      (* Pneomatic ->  FB_Piston *)
'2AAx001',   'Error',   'Waiting for Sensor Open at Open command',
'2AAx002',   'Error',   'Waiting for Sensor NotClose at Open command',
'2AAx003',   'Error',   'Waiting for Sensor Close at Close command',
'2AAx004',   'Error',   'Waiting for Sensor NotOpen at Close command',
'2AAx005',   'Error',   'No Status',
'2AAx006',   'Error',   'No Valve Operation',
'2AAx007',   'Error',   'Not synchronized with last auto-cycle command',
'2AAx008',   'Error',   'Sensors Checking',	 
		(*Process elementts*)
'109x000x001',   'Warning',   'Conveyor 5 is full',
'109x000x002',   'Error',     'Conveyor 5 is full and Conveyor 4 is ready to output full stack',

'109x000x003',   'Warning',   'Slices Stack is Too Light',
'109x000x004',   'Error',     'Slices Stack is Too Light',

'109x000x005',   'Warning',   'Slices Stack is Too Heavy',
'109x000x006',   'Error',     'Slices Stack is Too Heavy',
 
'555x000x001',   'Error',     'Hello world from NIV',

'985x000x001',   'Warning',     'X lens Constant velocity did not reach during coating',



(*Niv Section*)
(*Cycle X Curtain*)
(*Cycle X & Y*)
(*Cycle X & Theta)
(*Nozzle Operation*)
(*Cycle X Curtain*)
(*Cycle X Curtain*)*)




''];		
END_VAR

// ---- 01 Instance/06-Visu/g_Common.TcGVL
{attribute 'qualified_only'}
VAR_GLOBAL
	iContent_Main: INT;

END_VAR

// ---- 01 Instance/07-Mode/GVL_OperMode.TcGVL
VAR_GLOBAL

	eLightTowerState: E_LightTowerState;
	eBuzzerMode: E_BuzzerMode;
	bBuzzerMute: BOOL;

	bPauseMachine: BOOL;
	bResumeMachine: BOOL;
	bResetAllCycles: BOOL;
	
	PauseAll: BOOL;
	PauseAllDelayed: BOOL;
	ResumeAll: BOOL;	

	iActErrors							: INT;
	iActMessages						: INT;
	iActWarning							: INT;

	fbMode	: ARRAY[0..E_ModeZone.eLast] OF FB_ModeSelect;
	stMode	: ARRAY[0..E_ModeZone.eLast] OF ST_Mode;
	stOper	: ARRAY[0..E_ModeZone.eLast] OF ST_OperationButtons;
	
	fbLightTower: ARRAY[0..E_SkidZone.eLast] OF FB_LightTower;
	fbLightTower_Control: ARRAY[0..E_SkidZone.eLast] OF FB_LightTower_Control;



	//Operational Modes	
	stModeMain: ST_Mode;
	
	// Operational Buttons
	stOpMain				:ST_OperationButtons;
	stOpNonPause			:ST_OperationButtons;	

END_VAR

// ---- 01 Instance/12 Analog Sensor/g_AnalogSensor.TcGVL
//{attribute 'qualified_only'}
VAR_GLOBAL	
	fbAnalogSensor			: ARRAY[0..E_ASense_Name.last] OF FB_AnalogSensor;
	
	//arAnalogSensorName		: ARRAY[0..E_ASense_Name.last] OF STRING(12);
	
	//arAnalogSensorRawValue	: ARRAY[0..E_ASense_Name.last] OF INT;

	iAnalogSensor_sel		: INT:=1;
	
	arAnalogSensorNameList	: ARRAY[0..E_ASense_Name.last] OF STRING(12);
	eAnalogSensorNameList	: E_ASense_Name;

	
END_VAR
//{attribute 'qualified_only'}
VAR_GLOBAL PERSISTENT
	//stAnalogSensorSetting	: ARRAY[0..E_Pis_Name.last] OF ST_Piston_Setting_Param;
	stAnalogSensor			: ARRAY[0..E_ASense_Name.last] OF ST_AnalogSensor;
END_VAR

VAR_GLOBAL CONSTANT

END_VAR

// ---- 01 Instance/13 Process Control/g_ProcControl.TcGVL
//{attribute 'qualified_only'}
VAR_GLOBAL
	//concentration
	(*stDetergent					:	ST_ProcessControl	;
	pcDetergent					: 	FB_ProcessControl	;	//detergent local
	stDisinfectant				:	ST_ProcessControl	;
	pcDisinfectant				: 	FB_ProcessControl	;	//detergent local
    //temperature
	stTemperature_Deterg			:	ST_ProcessControl	;
	pcTemperature_Deterg			: 	FB_ProcessControl	;	//detergent Client	
	stTemperature_Dis				:	ST_ProcessControl	;
	pcTemperature_Dis				: 	FB_ProcessControl	;//disinfectant local/client
	
	//flow rate
	stFlow_Rate						:	ST_ProcessControl	;//CIP
	pcFlow_Rate						: 	FB_ProcessControl	;//disinfectant local/client
	stFlow_Rate_2					:	ST_ProcessControl	;//CLient CIP //level control 
	pcFlow_Rate_2					: 	FB_ProcessControl	;//disinfectant local/client //level control 
	
	//colar marinade 
	//pressure
	stPressure						:	ST_ProcessControl	;
	pcPressure						: 	FB_ProcessControl	;//CIP //Client	
	*)
	
	///////////////////ARRAYS///////////////////
	arr_fbProcCntrl			:	ARRAY [0..E_ProcessControl_Name.eProcCntrl_Last] OF FB_ProcessControl	;
	arr_ProcCntrl_NameList	:	ARRAY [0..E_ProcessControl_Name.eProcCntrl_Last] OF STRING	;
	eProcCntrl_Name			: E_ProcessControl_Name;
END_VAR
VAR_GLOBAL PERSISTENT
	arr_stProcCntrl			:	ARRAY [0..E_ProcessControl_Name.eProcCntrl_Last] OF ST_ProcessControl	;
END_VAR

// ---- 03 Project/12 TriBlender/g_HMI_Panel.TcGVL
//{attribute 'qualified_only'}
VAR_GLOBAL
	stVisuPLC_To_PLC		AT %MB1000 : ST_VisuPLC_To_PLC;
	stPLC_To_VisuPLC		AT %MB2000 : ST_PLC_To_VisuPLC;
	
	i_stVisuPLC_To_PLC		AT %I* : ST_VisuPLC_To_PLC;
	q_stPLC_To_VisuPLC		AT %Q* : ST_PLC_To_VisuPLC;	
END_VAR

// ---- 03 Project/15 Production Recipes/g_Prod.TcGVL
{attribute 'qualified_only'}
VAR_GLOBAL PERSISTENT
	
	arrRecipeMarinade	: ARRAY[1..cMax_Prod_Recipe] OF ST_Prod_Recipe;
	arrRecipeColor		: ARRAY[1..cMax_Prod_Recipe] OF ST_Prod_Recipe;
	
	iUserSelected_Marinade	: INT;
	iUserSelected_Color		: INT;
	
	fbProdRecipe_Manage	: FB_ProdRecipe_Manage;
	
	listRecipe_Marinade	: ARRAY[1..cMax_Prod_Recipe] OF STRING(30);
	listRecipe_Color	: ARRAY[1..cMax_Prod_Recipe] OF STRING(30);
	
	dtProdTimePicker	: DATE_AND_TIME;
	dtProdTimeMin		: DATE_AND_TIME;
	dtProdTimeMax		: DATE_AND_TIME;



END_VAR
VAR_GLOBAL CONSTANT 
	cMax_Prod_Recipe	: INT:=10;
	cMaxCompInProduct	: USINT:= 10;
END_VAR

// ---- 03 Project/30 IO/gIO.TcGVL
//{attribute 'qualified_only'}
VAR_GLOBAL
	i_EL			AT %I*	: ARRAY[1..27] 		OF ST_EL18x9;
	q_EL			AT %Q*	: ARRAY[1..11] 		OF ST_EL28x9;
	ai_EL			AT %I*	: ARRAY[1..6] 		OF ST_EL3xx8;
	aq_EL			AT %Q*	: ARRAY[1..1] 		OF ST_EL4xx8;

	
	q_Manifold1 	AT %Q*	: ARRAY[1..24] 		OF ST_VTUG;
	q_Manifold2 	AT %Q*	: ARRAY[1..24] 		OF ST_VTUG;
	q_Manifold3 	AT %Q*	: ARRAY[1..24] 		OF ST_VTUG;

	Nidec					: ARRAY[0..E_Pump_List.last] 		OF ST_Nidec;

	
	arSafe			: ARRAY[1..1] OF ST_TwinSAFE;
	bStateSafe		: BOOL;
	bStateSafe_ES1	: BOOL;
	bStateSafe_ES2	: BOOL;
	bStateSafe_ES3	: BOOL;
	bStateSafe_ES4	: BOOL;
	
	fbScaleFactor: ARRAY[0..E_ASense_Name.last] 		OF FB_ScaleFactor;

	
END_VAR

// ---- 03 Project/g_Data.TcGVL
//{attribute 'qualified_only'}
VAR_GLOBAL PERSISTENT
	gCIP_ValvUL			:	ARRAY [1..8,1..6] OF E_Pis_Name	:=[
																E_Pis_Name.V3004,E_Pis_Name.V3017,E_Pis_Name.V3023,E_Pis_Name.e0_not_in_use,E_Pis_Name.e0_not_in_use,E_Pis_Name.e0_not_in_use,
																E_Pis_Name.V3010,E_Pis_Name.V3027,E_Pis_Name.V3028,E_Pis_Name.e0_not_in_use,E_Pis_Name.e0_not_in_use,E_Pis_Name.e0_not_in_use,
																E_Pis_Name.V4034,E_Pis_Name.V4004,E_Pis_Name.V4017,E_Pis_Name.v4023,E_Pis_Name.e0_not_in_use,E_Pis_Name.e0_not_in_use,
																E_Pis_Name.V4033,E_Pis_Name.V4010,E_Pis_Name.V4027,E_Pis_Name.V4028,E_Pis_Name.e0_not_in_use,E_Pis_Name.e0_not_in_use,
																
																E_Pis_Name.V3113,E_Pis_Name.V3004,E_Pis_Name.V3010,E_Pis_Name.V3023,E_Pis_Name.V3028,E_Pis_Name.e0_not_in_use,
																E_Pis_Name.v2114,E_Pis_Name.V4004,E_Pis_Name.V4010,E_Pis_Name.V2116,E_Pis_Name.V4023,E_Pis_Name.V4028,
																E_Pis_Name.V3017,E_Pis_Name.V3027,E_Pis_Name.e0_not_in_use,E_Pis_Name.e0_not_in_use,E_Pis_Name.e0_not_in_use,E_Pis_Name.e0_not_in_use,
																E_Pis_Name.V4017,E_Pis_Name.v4027,E_Pis_Name.V2115,E_Pis_Name.V4034,E_Pis_Name.V4033,E_Pis_Name.e0_not_in_use														
															];	
	gCIP_ValvUL_Seat	:	ARRAY [1..8,1..6] OF BOOL :=[
															0,1,1,0,0,0, // Client 1 eTank_1,
															0,1,1,0,0,0, // Client 2 eTank_2,
															0,0,1,1,0,0, // Client 3 eTank_3,
															0,0,1,1,0,0, // Client 4 eTank_4,
															0,1,1,0,0,0, // Client 5
															0,1,1,0,0,0, // Client 6
															0,0,0,0,0,0, // Client 7
															0,0,0,1,1,0 // Client 8 
														]	;	//0-Low, 1-Up

	fbElement: ARRAY[1..8] OF FB_Element;
	
	fbIntCon_TriB_T1_Marin	: FB_InterConnection;
	fbIntCon_TriB_T2_Marin	: FB_InterConnection;
	fbIntCon_TriB_T3_Color	: FB_InterConnection;
	fbIntCon_TriB_T4_Color	: FB_InterConnection;
	fbIntCon_ProL_T1_Marin	: FB_InterConnection;
	fbIntCon_ProL_T2_Marin	: FB_InterConnection;
	fbIntCon_ProL_T3_Color	: FB_InterConnection;
	fbIntCon_ProL_T4_Color	: FB_InterConnection;
	
	fbTank1					: FB_ProductionTank;
	fbTank2					: FB_ProductionTank;
	fbTank3					: FB_ProductionTank;
	fbTank4					: FB_ProductionTank;

	fbTankTarget_1				: FB_Tank_Target;
	fbTankTarget_2				: FB_Tank_Target;
	fbTankTarget_3				: FB_Tank_Target;
	fbTankTarget_4				: FB_Tank_Target;

	fbLineSource_Marinade		: FB_Line_Source;
	fbTriBlenderSource_Marinade	: FB_Line_Source;
	fbLineSource_Color			: FB_Line_Source;
	fbTriBlenderSource_Color	: FB_Line_Source;
	
	fbLineTarget_Marinade		: FB_Line_Target;
	fbTriBlenderTarget_Marinade	: FB_Line_Target;
	fbLineTarget_Color			: FB_Line_Target;
	fbTriBlenderTarget_Color	: FB_Line_Target;
	
	fbCIP						: FB_CIP;
	
	fbCIP_Source				: FB_CIP_Source;
	fbCIP_Return				: FB_CIP_Return;
	fbCIP_Client				: FB_CIP_Client;
	
	fbCIP_ClientTank_Marinade	: FB_CIP_ClientTank;
	fbCIP_ClientTank_Color		: FB_CIP_ClientTank;

	fbDissolving				: FB_Dissolving;
	fbTriBlender_Select			: FB_TriBlender_Select;
	eTriBlenderUsage	: E_TriBlenderUsage;
	
	eTriBlenderPipe		: E_TriBlenderPipe;
	eTriBlenderPipe_In	: E_TriBlenderPipe;
	eTriBlenderPipe_Out	: E_TriBlenderPipe;

	ePrL_M_Usage		: E_PrLine_M_LineUsage;
	ePrL_C_Usage		: E_PrLine_C_Usage;
	
	//Pumps
	//fbPumpLine_P4001		:	FB_Pump	;
	//fbPumpLine_P3001		:	FB_Pump	;
	//fbPumpTriblender_TB001	:	FB_Pump	;
	
	arCIP_RequestBufer: ARRAY [0..9] OF ST_CIP_Request;

	//stDev			: 	ARRAY[0..E_OwnerDevice.common] OF 	ST_DeviceErrorHandeling;
	//stDev			: 	ARRAY[0..E_OwnerDevice.common] OF 	ST_OperationButtons;
	
	//Valves
	arr_TankValves					:	ARRAY [1..4] OF st_TankValves		;
	arr_LineSourceValves			:	ARRAY [1..4] OF st_LineSourceValves	;
	arr_TriBlenderSourceValves		:	ARRAY [1..4] OF st_LineSourceValves	;
	arr_LineTargetValves			:	ARRAY [1..4] OF st_LineTargetValves	;
	arr_fbTriBlenderTargetValves	:	ARRAY [1..4] OF st_LineTargetValves	;
	
	//Sensors
	(*lvl_Tank_T91	: ST_Tank_Level	;
	lvl_Tank_T92	: ST_Tank_Level	;
	lvl_Tank_T93	: ST_Tank_Level	;
	lvl_Tank_T94	: ST_Tank_Level	;
	
	lvl_Tank_T91_Analog	:	ST_AnalogSignal	;
	lvl_Tank_T92_Analog	:	ST_AnalogSignal	;
	lvl_Tank_T93_Analog	:	ST_AnalogSignal	;
	lvl_Tank_T94_Analog	:	ST_AnalogSignal	;
	
	fbLvl_Tank_T91	:	FB_TankLevel	;
	fbLvl_Tank_T92	:	FB_TankLevel	;
	fbLvl_Tank_T93	:	FB_TankLevel	;
	fbLvl_Tank_T94	:	FB_TankLevel	;
	
	fb_Tank_T91_Sensors	:	FB_TankSensors	;
	fb_Tank_T92_Sensors	:	FB_TankSensors	;
	fb_Tank_T93_Sensors	:	FB_TankSensors	;
	fb_Tank_T94_Sensors	:	FB_TankSensors	;*)
	
	//Heat Exchanger
	fbHeatExchenger	:	FB_HeatExchanger	;
	stHeatExchanger	:	ST_HeatExchanger	;
	
	////////////////////////////////////////////////////////////////
	arrTanksSens	:	ARRAY [0..E_Tank_Name.last] OF FB_TankSensors;
	stTanksSens		:	ARRAY [0..E_Tank_Name.last] OF ST_Tank_Level;
	
	////////////////////////////////////////////////////////////////
	arr_CIP_Param		:	ARRAY [0..E_CIP_Usage.eLocal] OF ST_CIP_Param		;//9-local, 1..8 cleints
	
	//additional variables
	b_CIP_Run	:	BOOL	;
	bDisolvingProcess_Active: BOOL;
	bDisolvingProcess_Done: BOOL;
	
	ExDuration_Default				: TIME:=T#48H;	//Expiration
	ExDuration_Default_Line			: TIME:=T#24H;	//Expiration
	ExDuration_Default_LineStandby	: TIME:=T#2H;	//Expiration

	//arr_ProdTank		:	ARRAY [0..E_Tank_Name.last] OF ST_ProdParams;
	
	//stTriBlender		: ST_TriBlender;		
	//arrProductionComponents	: ARRAY [0..g_Prod.cMaxCompInProduct-1] OF ST_Component;
END_VAR
VAR_GLOBAL CONSTANT
	
END_VAR

// ---- 00 Library/03 SFC/ITF_FB_SFC_Cycle.TcIO
INTERFACE ITF_FB_SFC_Cycle

METHOD m_Set_SFCFlags_Reference : BOOL
VAR_INPUT
END_VAR
END_METHOD

END_INTERFACE

// ---- 01 Instance/04 Recipe/prg_Call_Recipe_Slow.TcPOU
PROGRAM prg_Call_Recipe_Slow
VAR
	i							: INT;
	bFirstScan					: BOOL:= TRUE;
	ton_RecipeReady				: TON;
	
	
	eRecipeName: E_Recipe_Name;

	r_trigAxisPoints_Loaded: R_TRIG;
	ton_WriteLoaded_Points: TON;
	r_trigRecipe3_loaded: R_TRIG;

	bAllRecipesLoaded: BOOL;
	iRecipeSwitchFrameVar: INT;
	bLoadDefForAll: BOOL;
	
	tPath: STRING(80);
END_VAR

act_Set_StoragePath_For_All();
//act_LoadDeafult();

ton_RecipeReady(PT:=T#1S, IN:=GVL_Recipe.stRecipe[1].bInit AND bFirstScan);
IF ton_RecipeReady.Q THEN;
	bFirstScan:=FALSE;
	bLoadDefForAll:=TRUE;
END_IF




(********************  Other Instances Recipes******************************) // 
FOR eRecipeName:=1 TO E_Recipe_Name.R_Piston_Settings DO	
	fbRecipe[eRecipeName](pstRecipe:=ADR(GVL_Recipe.stRecipe[eRecipeName]), 
			bMemoRecipeUpdated:=, 
			sRecipeDef:=TO_STRING(eRecipeName),
			bLoadDefault:=ar_RecipesLoadDefault[eRecipeName],
			bHMI_FrameActive:=iRecipeSwitchFrameVar=eRecipeName-1,//changed
			sRecipesStoragePath:=ar_RecipesStoragePath[eRecipeName]);
END_FOR
(*			
IF (*fbRecipe_1.bMemoRecipeUpdated AND*) 
fbRecipe_2.bMemoRecipeUpdated 
AND fbRecipe_3.bMemoRecipeUpdated 
AND fbRecipe_4.bMemoRecipeUpdated 
AND fbRecipe_5.bMemoRecipeUpdated 
THEN;
	bAllRecipesLoaded:=TRUE;
ELSE;
	bAllRecipesLoaded:=FALSE;
END_IF
*)

ACTION act_LoadDeafult:
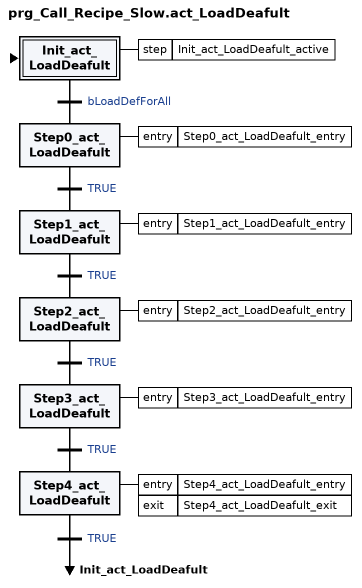
INITIAL_STEP Init_act_LoadDeafult:
    Init_act_LoadDeafult_active(N);  // step action
END_STEP
TRANSITION FROM Init_act_LoadDeafult TO Step0_act_LoadDeafult
    := bLoadDefForAll;
END_TRANSITION
STEP Step0_act_LoadDeafult:  // min time T#2s
    Step0_act_LoadDeafult_entry(P1);  // entry action
END_STEP
TRANSITION FROM Step0_act_LoadDeafult TO Step1_act_LoadDeafult
    := TRUE;
END_TRANSITION
STEP Step1_act_LoadDeafult:  // min time T#2s
    Step1_act_LoadDeafult_entry(P1);  // entry action
END_STEP
TRANSITION FROM Step1_act_LoadDeafult TO Step2_act_LoadDeafult
    := TRUE;
END_TRANSITION
STEP Step2_act_LoadDeafult:  // min time T#2s
    Step2_act_LoadDeafult_entry(P1);  // entry action
END_STEP
TRANSITION FROM Step2_act_LoadDeafult TO Step3_act_LoadDeafult
    := TRUE;
END_TRANSITION
STEP Step3_act_LoadDeafult:  // min time T#2s
    Step3_act_LoadDeafult_entry(P1);  // entry action
END_STEP
TRANSITION FROM Step3_act_LoadDeafult TO Step4_act_LoadDeafult
    := TRUE;
END_TRANSITION
STEP Step4_act_LoadDeafult:  // min time T#2s
    Step4_act_LoadDeafult_entry(P1);  // entry action
    Step4_act_LoadDeafult_exit(P0);  // exit action
END_STEP
TRANSITION FROM Step4_act_LoadDeafult TO Init_act_LoadDeafult
    := TRUE;
END_TRANSITION
END_ACTION

ACTION act_Set_StoragePath_For_All:
FOR eRecipeName:=1 TO E_Recipe_Name.R_Piston_Settings DO;
	GVL_Recipe.ar_RecipesStoragePath_Folder[eRecipeName]:=TO_STRING(eRecipeName);
	tPath:='';
	tPath:=CONCAT(tPath,GVL_Recipe.ar_RecipesStoragePath_Root[GVL_Recipe.eRecipeRootFolder]);
	tPath:=CONCAT(tPath,'\');
	tPath:=CONCAT(tPath,TO_STRING(eRecipeName));
	tPath:=CONCAT(tPath,'\');
	GVL_Recipe.ar_RecipesStoragePath[eRecipeName]:=tPath;
(*
	GVL_Recipe.ar_RecipesStoragePath[eRecipeName]:=
			CONCAT(	GVL_Recipe.ar_RecipesStoragePath_Root[GVL_Recipe.eRecipeRootFolder],'\'); 
	GVL_Recipe.ar_RecipesStoragePath[eRecipeName]:=		
			CONCAT(	GVL_Recipe.ar_RecipesStoragePath[eRecipeName],TO_STRING(eRecipeName));
	GVL_Recipe.ar_RecipesStoragePath[eRecipeName]:=		
			CONCAT(	GVL_Recipe.ar_RecipesStoragePath[eRecipeName],'1');				
	GVL_Recipe.ar_RecipesStoragePath[eRecipeName]:=		
			CONCAT(	GVL_Recipe.ar_RecipesStoragePath[eRecipeName],'\');		
*)	
END_FOR
END_ACTION

ACTION Init_act_LoadDeafult_active:
GVL_Recipe.ar_RecipesLoadDefault[1]:=FALSE;
GVL_Recipe.ar_RecipesLoadDefault[2]:=FALSE;
GVL_Recipe.ar_RecipesLoadDefault[3]:=FALSE;
GVL_Recipe.ar_RecipesLoadDefault[4]:=FALSE;
GVL_Recipe.ar_RecipesLoadDefault[5]:=FALSE;
END_ACTION

ACTION Step0_act_LoadDeafult_entry:
GVL_Recipe.ar_RecipesLoadDefault[1]:=TRUE;
END_ACTION

ACTION Step1_act_LoadDeafult_entry:
GVL_Recipe.ar_RecipesLoadDefault[2]:=TRUE;
END_ACTION

ACTION Step2_act_LoadDeafult_entry:
GVL_Recipe.ar_RecipesLoadDefault[3]:=TRUE;
END_ACTION

ACTION Step3_act_LoadDeafult_entry:
GVL_Recipe.ar_RecipesLoadDefault[4]:=TRUE;
END_ACTION

ACTION Step4_act_LoadDeafult_entry:
GVL_Recipe.ar_RecipesLoadDefault[5]:=TRUE;
END_ACTION

ACTION Step4_act_LoadDeafult_exit:
bLoadDefForAll:=FALSE;
END_ACTION

END_PROGRAM

// ---- POUs/MAIN.TcPOU
PROGRAM MAIN
VAR

	fTotalCIP_Volume: REAL;
	fbWritePersistent: FB_WritePersistentData;
	bTesting		:	BOOL:=FALSE	;
	nI_1			: 	INT		;
	ftg_EStop_Fall	: 	F_TRIG	;
	rs_EStopFall	: 	RS	;
	bTestEstop		:	BOOL:=TRUE	;
	FB_OpenClose_Vlave_4026: FB_OpenClose_Vlave;
	bTemp_Water_Overweight_check: BOOL;
	fbUPS: FB_S_UPS_CX51x0;

	bSetExpeationTime: BOOL;
	i: E_ELEMENT_LIST;
	tExpirationSet_Test: TIME := T#10s;
END_VAR

prg_RealClock();
prg_Piston();
prg_Safety();
prg_MessageManager();
prg_Messages();
prg_Call_OpMode();
prg_IntCheck();
prg_User();
act_ResetPumps();
(*
prg_TriBlender(
		fb_TriBlenderPump:= g_Pump.fbPump[E_Pump_List.TB0001],
		stTriblender:=stTriblender,
		arrComponents:=arrProductionComponents);
*)		
//act_SetAnalogSens_Test();//To be deleted, for testing purposes
act_Call_Sensors_Analog();//To be deleted, for testing purposes
act_Call_Sensors_Analog_1();//To be deleted, for testing purposes
act_Call_ScaleFactor();//To be deleted, for testing purposes
act_Call_ProcessCntrl();

act_SetValves();
act_ClientPump_Select();
act_ClientStirrer_Select();
act_Call_Elements();
act_Call_Elements_Imp();
act_Call_Pumps();
prg_InterCon_Usage();
act_Sensors();
act_HeatExchenger();
act_Call_CIP();
act_Call_Production();

act_Call_For_HMI();

g_SFC.fbSFC_Temp1();

//Temtprary Overweght protection!!!!! DO NOT DELETE
IF fTotalCIP_Volume >=1500 AND FALSE THEN;
	//fbPis[E_Pis_Name.V1022].m_SetByRecipe(stPis:=stPis[E_Pis_Name.V1022], req:=E_Piston_Recipe_State.Release);
	//fbPis[E_Pis_Name.V1019].m_SetByRecipe(stPis:=stPis[E_Pis_Name.V1019], req:=E_Piston_Recipe_State.Release);
	//fbPis[E_Pis_Name.V1016].m_SetByRecipe(stPis:=stPis[E_Pis_Name.V1016], req:=E_Piston_Recipe_State.Release);
	//fbPis[E_Pis_Name.V1011].m_SetByRecipe(stPis:=stPis[E_Pis_Name.V1011], req:=E_Piston_Recipe_State.Release);
	bTemp_Water_Overweight_check:=FALSE;
	fbPrintErrMessageByID(sModuleDescription:='CIP',sActErrorID:='101x000x000');
ELSIF fTotalCIP_Volume < 1480 THEN;
	bTemp_Water_Overweight_check:=TRUE;
END_IF

IF arrTanksSens[E_Tank_Name.T91].get_stTankLevel_OverFlow() THEN;
	fbPis[E_Pis_Name.V1022].m_SetByRecipe(stPis:=stPis[E_Pis_Name.V1022], req:=E_Piston_Recipe_State.Release);
	//print error
	fbPrintErrMessageByID(sModuleDescription:='CIP',sActErrorID:='101x000x001');		
END_IF
IF arrTanksSens[E_Tank_Name.T92].get_stTankLevel_OverFlow() THEN;
	fbPis[E_Pis_Name.V1019].m_SetByRecipe(stPis:=stPis[E_Pis_Name.V1019], req:=E_Piston_Recipe_State.Release);
	//print error
	fbPrintErrMessageByID(sModuleDescription:='CIP',sActErrorID:='101x000x002');		
END_IF
IF arrTanksSens[E_Tank_Name.T93].get_stTankLevel_OverFlow() THEN;
	fbPis[E_Pis_Name.V1016].m_SetByRecipe(stPis:=stPis[E_Pis_Name.V1016], req:=E_Piston_Recipe_State.Release);
	//print error	
	fbPrintErrMessageByID(sModuleDescription:='CIP',sActErrorID:='101x000x003');	
END_IF
IF arrTanksSens[E_Tank_Name.T94].get_stTankLevel_OverFlow() THEN;
	fbPis[E_Pis_Name.V1011].m_SetByRecipe(stPis:=stPis[E_Pis_Name.V1011], req:=E_Piston_Recipe_State.Release);
	//print error
	fbPrintErrMessageByID(sModuleDescription:='CIP',sActErrorID:='101x000x004');		
END_IF
	
IF bSetExpeationTime THEN;
	bSetExpeationTime:=FALSE;
	FOR i:=E_Element_List.eTank_1 TO E_Element_List.eLine_Color DO
		fbElement[i].ExpirationTime:=tExpirationSet_Test;
		
	END_FOR
END_IF
	

mElementList_SetName();

fbWritePersistent(
	NETID:= , 
	PORT:= 851, 
	START:= , 
	TMOUT:= T#3S, 
	MODE:= , 
	BUSY=> , 
	ERR=> , 
	ERRID=> );

fbUPS();

ACTION act_Call_CIP:
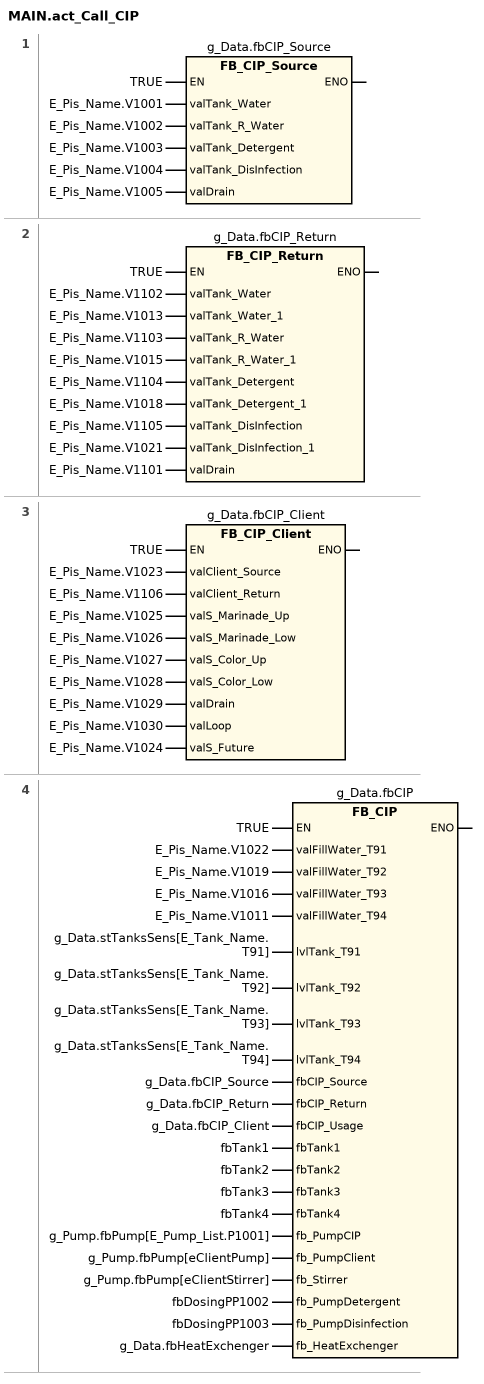
// NETWORK 1
g_Data.fbCIP_Source(
    valTank_Water := E_Pis_Name.V1001,
    valTank_R_Water := E_Pis_Name.V1002,
    valTank_Detergent := E_Pis_Name.V1003,
    valTank_DisInfection := E_Pis_Name.V1004,
    valDrain := E_Pis_Name.V1005); // FB_CIP_Source

// NETWORK 2
g_Data.fbCIP_Return(
    valTank_Water := E_Pis_Name.V1102,
    valTank_Water_1 := E_Pis_Name.V1013,
    valTank_R_Water := E_Pis_Name.V1103,
    valTank_R_Water_1 := E_Pis_Name.V1015,
    valTank_Detergent := E_Pis_Name.V1104,
    valTank_Detergent_1 := E_Pis_Name.V1018,
    valTank_DisInfection := E_Pis_Name.V1105,
    valTank_DisInfection_1 := E_Pis_Name.V1021,
    valDrain := E_Pis_Name.V1101); // FB_CIP_Return

// NETWORK 3
g_Data.fbCIP_Client(
    valClient_Source := E_Pis_Name.V1023,
    valClient_Return := E_Pis_Name.V1106,
    valS_Marinade_Up := E_Pis_Name.V1025,
    valS_Marinade_Low := E_Pis_Name.V1026,
    valS_Color_Up := E_Pis_Name.V1027,
    valS_Color_Low := E_Pis_Name.V1028,
    valDrain := E_Pis_Name.V1029,
    valLoop := E_Pis_Name.V1030,
    valS_Future := E_Pis_Name.V1024); // FB_CIP_Client

// NETWORK 4
g_Data.fbCIP(
    valFillWater_T91 := E_Pis_Name.V1022,
    valFillWater_T92 := E_Pis_Name.V1019,
    valFillWater_T93 := E_Pis_Name.V1016,
    valFillWater_T94 := E_Pis_Name.V1011,
    lvlTank_T91 := g_Data.stTanksSens[E_Tank_Name.T91],
    lvlTank_T92 := g_Data.stTanksSens[E_Tank_Name.T92],
    lvlTank_T93 := g_Data.stTanksSens[E_Tank_Name.T93],
    lvlTank_T94 := g_Data.stTanksSens[E_Tank_Name.T94],
    fbCIP_Source := g_Data.fbCIP_Source,
    fbCIP_Return := g_Data.fbCIP_Return,
    fbCIP_Usage := g_Data.fbCIP_Client,
    fbTank1 := fbTank1,
    fbTank2 := fbTank2,
    fbTank3 := fbTank3,
    fbTank4 := fbTank4,
    fb_PumpCIP := g_Pump.fbPump[E_Pump_List.P1001],
    fb_PumpClient := g_Pump.fbPump[eClientPump],
    fb_Stirrer := g_Pump.fbPump[eClientStirrer],
    fb_PumpDetergent := fbDosingPP1002,
    fb_PumpDisinfection := fbDosingPP1003,
    fb_HeatExchenger := g_Data.fbHeatExchenger); // FB_CIP

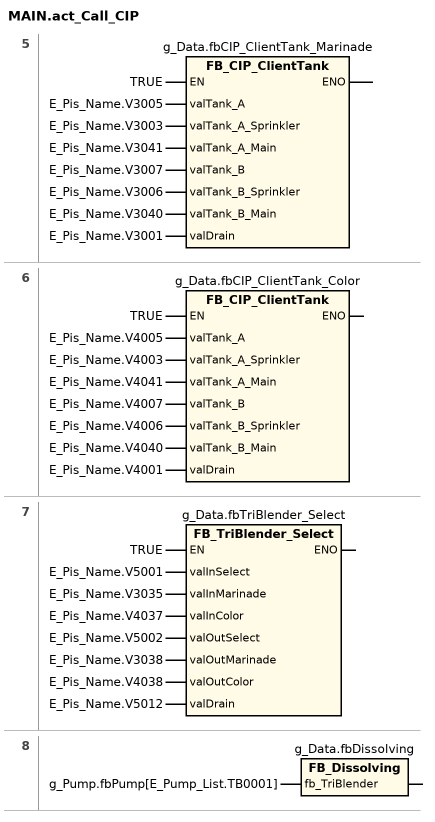
// NETWORK 5
g_Data.fbCIP_ClientTank_Marinade(
    valTank_A := E_Pis_Name.V3005,
    valTank_A_Sprinkler := E_Pis_Name.V3003,
    valTank_A_Main := E_Pis_Name.V3041,
    valTank_B := E_Pis_Name.V3007,
    valTank_B_Sprinkler := E_Pis_Name.V3006,
    valTank_B_Main := E_Pis_Name.V3040,
    valDrain := E_Pis_Name.V3001); // FB_CIP_ClientTank

// NETWORK 6
g_Data.fbCIP_ClientTank_Color(
    valTank_A := E_Pis_Name.V4005,
    valTank_A_Sprinkler := E_Pis_Name.V4003,
    valTank_A_Main := E_Pis_Name.V4041,
    valTank_B := E_Pis_Name.V4007,
    valTank_B_Sprinkler := E_Pis_Name.V4006,
    valTank_B_Main := E_Pis_Name.V4040,
    valDrain := E_Pis_Name.V4001); // FB_CIP_ClientTank

// NETWORK 7
g_Data.fbTriBlender_Select(
    valInSelect := E_Pis_Name.V5001,
    valInMarinade := E_Pis_Name.V3035,
    valInColor := E_Pis_Name.V4037,
    valOutSelect := E_Pis_Name.V5002,
    valOutMarinade := E_Pis_Name.V3038,
    valOutColor := E_Pis_Name.V4038,
    valDrain := E_Pis_Name.V5012); // FB_TriBlender_Select

// NETWORK 8
g_Data.fbDissolving(fb_TriBlender := g_Pump.fbPump[E_Pump_List.TB0001]); // FB_Dissolving
END_ACTION

ACTION act_Call_Elements:
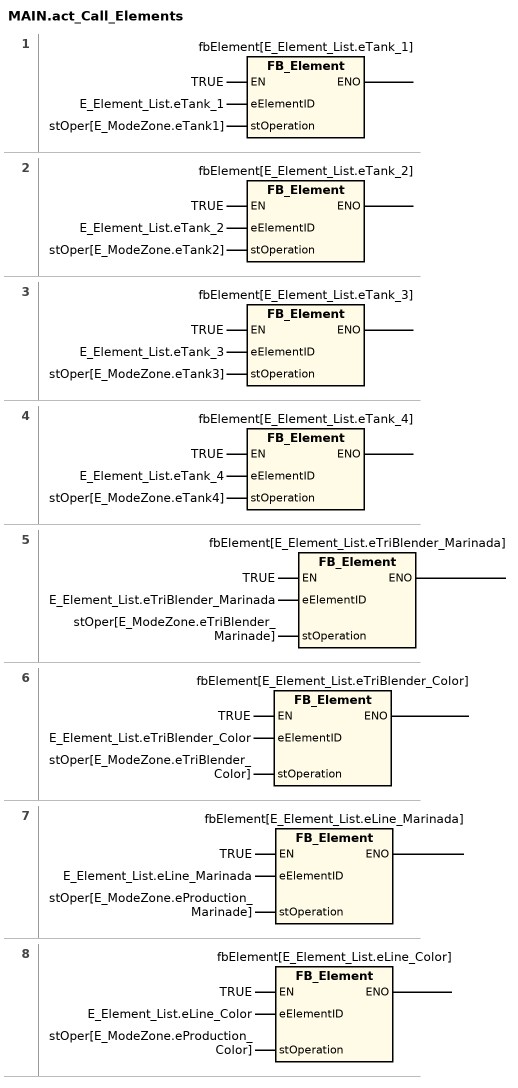
// NETWORK 1
fbElement[E_Element_List.eTank_1](eElementID := E_Element_List.eTank_1, stOperation := stOper[E_ModeZone.eTank1]); // FB_Element

// NETWORK 2
fbElement[E_Element_List.eTank_2](eElementID := E_Element_List.eTank_2, stOperation := stOper[E_ModeZone.eTank2]); // FB_Element

// NETWORK 3
fbElement[E_Element_List.eTank_3](eElementID := E_Element_List.eTank_3, stOperation := stOper[E_ModeZone.eTank3]); // FB_Element

// NETWORK 4
fbElement[E_Element_List.eTank_4](eElementID := E_Element_List.eTank_4, stOperation := stOper[E_ModeZone.eTank4]); // FB_Element

// NETWORK 5
fbElement[E_Element_List.eTriBlender_Marinada](eElementID := E_Element_List.eTriBlender_Marinada, stOperation := stOper[E_ModeZone.eTriBlender_Marinade]); // FB_Element

// NETWORK 6
fbElement[E_Element_List.eTriBlender_Color](eElementID := E_Element_List.eTriBlender_Color, stOperation := stOper[E_ModeZone.eTriBlender_Color]); // FB_Element

// NETWORK 7
fbElement[E_Element_List.eLine_Marinada](eElementID := E_Element_List.eLine_Marinada, stOperation := stOper[E_ModeZone.eProduction_Marinade]); // FB_Element

// NETWORK 8
fbElement[E_Element_List.eLine_Color](eElementID := E_Element_List.eLine_Color, stOperation := stOper[E_ModeZone.eProduction_Color]); // FB_Element
END_ACTION

ACTION act_Call_Elements_Imp:
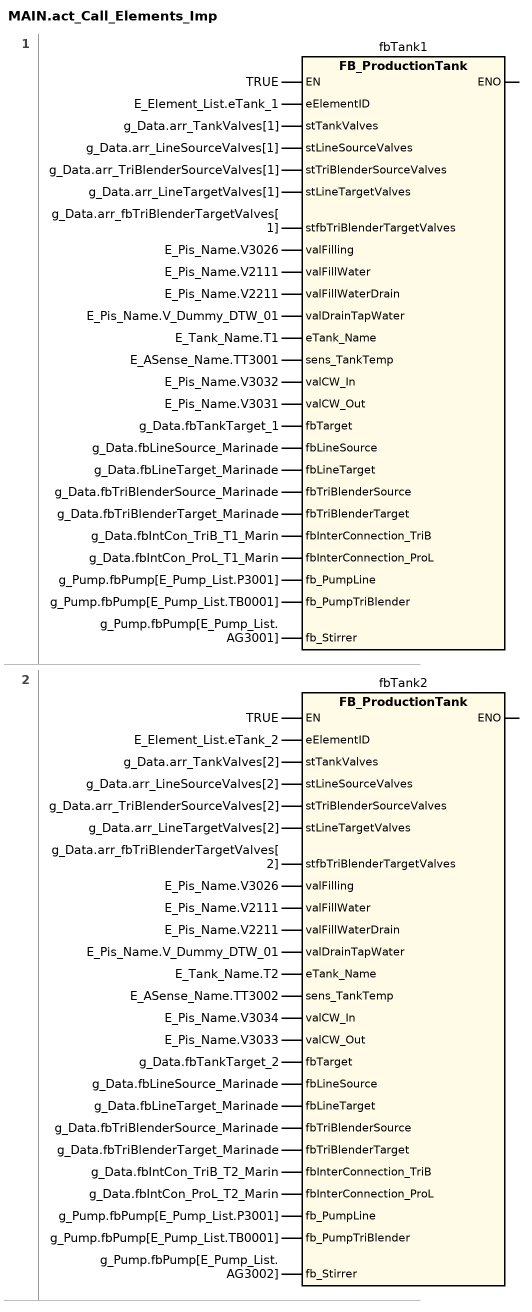
// NETWORK 1
fbTank1(
    eElementID := E_Element_List.eTank_1,
    stTankValves := g_Data.arr_TankValves[1],
    stLineSourceValves := g_Data.arr_LineSourceValves[1],
    stTriBlenderSourceValves := g_Data.arr_TriBlenderSourceValves[1],
    stLineTargetValves := g_Data.arr_LineTargetValves[1],
    stfbTriBlenderTargetValves := g_Data.arr_fbTriBlenderTargetValves[1],
    valFilling := E_Pis_Name.V3026,
    valFillWater := E_Pis_Name.V2111,
    valFillWaterDrain := E_Pis_Name.V2211,
    valDrainTapWater := E_Pis_Name.V_Dummy_DTW_01,
    eTank_Name := E_Tank_Name.T1,
    sens_TankTemp := E_ASense_Name.TT3001,
    valCW_In := E_Pis_Name.V3032,
    valCW_Out := E_Pis_Name.V3031,
    fbTarget := g_Data.fbTankTarget_1,
    fbLineSource := g_Data.fbLineSource_Marinade,
    fbLineTarget := g_Data.fbLineTarget_Marinade,
    fbTriBlenderSource := g_Data.fbTriBlenderSource_Marinade,
    fbTriBlenderTarget := g_Data.fbTriBlenderTarget_Marinade,
    fbInterConnection_TriB := g_Data.fbIntCon_TriB_T1_Marin,
    fbInterConnection_ProL := g_Data.fbIntCon_ProL_T1_Marin,
    fb_PumpLine := g_Pump.fbPump[E_Pump_List.P3001],
    fb_PumpTriBlender := g_Pump.fbPump[E_Pump_List.TB0001],
    fb_Stirrer := g_Pump.fbPump[E_Pump_List.AG3001]); // FB_ProductionTank

// NETWORK 2
fbTank2(
    eElementID := E_Element_List.eTank_2,
    stTankValves := g_Data.arr_TankValves[2],
    stLineSourceValves := g_Data.arr_LineSourceValves[2],
    stTriBlenderSourceValves := g_Data.arr_TriBlenderSourceValves[2],
    stLineTargetValves := g_Data.arr_LineTargetValves[2],
    stfbTriBlenderTargetValves := g_Data.arr_fbTriBlenderTargetValves[2],
    valFilling := E_Pis_Name.V3026,
    valFillWater := E_Pis_Name.V2111,
    valFillWaterDrain := E_Pis_Name.V2211,
    valDrainTapWater := E_Pis_Name.V_Dummy_DTW_01,
    eTank_Name := E_Tank_Name.T2,
    sens_TankTemp := E_ASense_Name.TT3002,
    valCW_In := E_Pis_Name.V3034,
    valCW_Out := E_Pis_Name.V3033,
    fbTarget := g_Data.fbTankTarget_2,
    fbLineSource := g_Data.fbLineSource_Marinade,
    fbLineTarget := g_Data.fbLineTarget_Marinade,
    fbTriBlenderSource := g_Data.fbTriBlenderSource_Marinade,
    fbTriBlenderTarget := g_Data.fbTriBlenderTarget_Marinade,
    fbInterConnection_TriB := g_Data.fbIntCon_TriB_T2_Marin,
    fbInterConnection_ProL := g_Data.fbIntCon_ProL_T2_Marin,
    fb_PumpLine := g_Pump.fbPump[E_Pump_List.P3001],
    fb_PumpTriBlender := g_Pump.fbPump[E_Pump_List.TB0001],
    fb_Stirrer := g_Pump.fbPump[E_Pump_List.AG3002]); // FB_ProductionTank

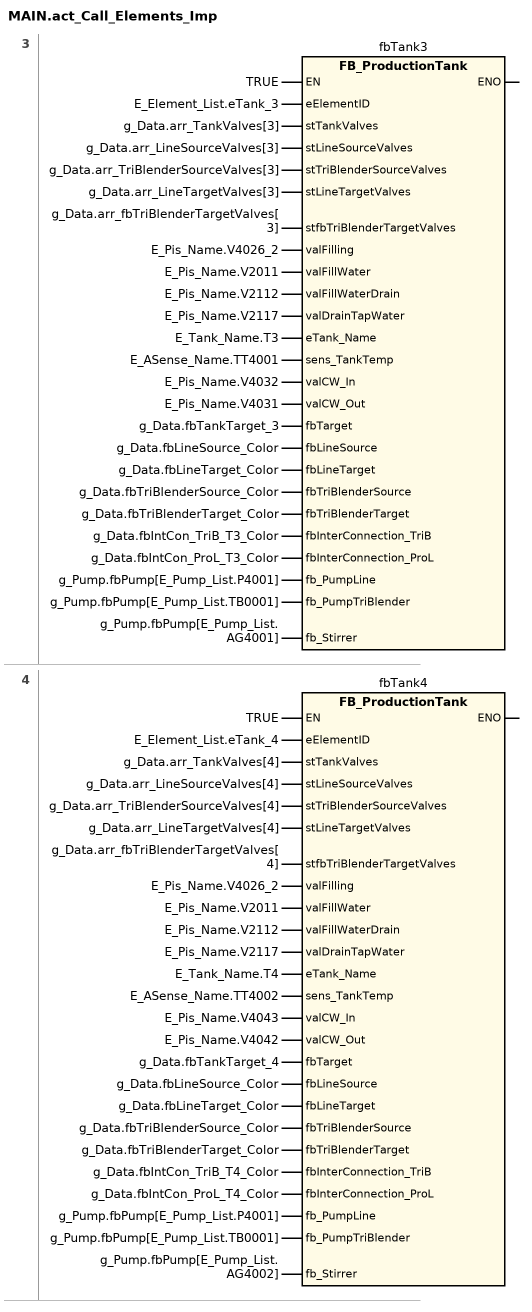
// NETWORK 3
fbTank3(
    eElementID := E_Element_List.eTank_3,
    stTankValves := g_Data.arr_TankValves[3],
    stLineSourceValves := g_Data.arr_LineSourceValves[3],
    stTriBlenderSourceValves := g_Data.arr_TriBlenderSourceValves[3],
    stLineTargetValves := g_Data.arr_LineTargetValves[3],
    stfbTriBlenderTargetValves := g_Data.arr_fbTriBlenderTargetValves[3],
    valFilling := E_Pis_Name.V4026_2,
    valFillWater := E_Pis_Name.V2011,
    valFillWaterDrain := E_Pis_Name.V2112,
    valDrainTapWater := E_Pis_Name.V2117,
    eTank_Name := E_Tank_Name.T3,
    sens_TankTemp := E_ASense_Name.TT4001,
    valCW_In := E_Pis_Name.V4032,
    valCW_Out := E_Pis_Name.V4031,
    fbTarget := g_Data.fbTankTarget_3,
    fbLineSource := g_Data.fbLineSource_Color,
    fbLineTarget := g_Data.fbLineTarget_Color,
    fbTriBlenderSource := g_Data.fbTriBlenderSource_Color,
    fbTriBlenderTarget := g_Data.fbTriBlenderTarget_Color,
    fbInterConnection_TriB := g_Data.fbIntCon_TriB_T3_Color,
    fbInterConnection_ProL := g_Data.fbIntCon_ProL_T3_Color,
    fb_PumpLine := g_Pump.fbPump[E_Pump_List.P4001],
    fb_PumpTriBlender := g_Pump.fbPump[E_Pump_List.TB0001],
    fb_Stirrer := g_Pump.fbPump[E_Pump_List.AG4001]); // FB_ProductionTank

// NETWORK 4
fbTank4(
    eElementID := E_Element_List.eTank_4,
    stTankValves := g_Data.arr_TankValves[4],
    stLineSourceValves := g_Data.arr_LineSourceValves[4],
    stTriBlenderSourceValves := g_Data.arr_TriBlenderSourceValves[4],
    stLineTargetValves := g_Data.arr_LineTargetValves[4],
    stfbTriBlenderTargetValves := g_Data.arr_fbTriBlenderTargetValves[4],
    valFilling := E_Pis_Name.V4026_2,
    valFillWater := E_Pis_Name.V2011,
    valFillWaterDrain := E_Pis_Name.V2112,
    valDrainTapWater := E_Pis_Name.V2117,
    eTank_Name := E_Tank_Name.T4,
    sens_TankTemp := E_ASense_Name.TT4002,
    valCW_In := E_Pis_Name.V4043,
    valCW_Out := E_Pis_Name.V4042,
    fbTarget := g_Data.fbTankTarget_4,
    fbLineSource := g_Data.fbLineSource_Color,
    fbLineTarget := g_Data.fbLineTarget_Color,
    fbTriBlenderSource := g_Data.fbTriBlenderSource_Color,
    fbTriBlenderTarget := g_Data.fbTriBlenderTarget_Color,
    fbInterConnection_TriB := g_Data.fbIntCon_TriB_T4_Color,
    fbInterConnection_ProL := g_Data.fbIntCon_ProL_T4_Color,
    fb_PumpLine := g_Pump.fbPump[E_Pump_List.P4001],
    fb_PumpTriBlender := g_Pump.fbPump[E_Pump_List.TB0001],
    fb_Stirrer := g_Pump.fbPump[E_Pump_List.AG4002]); // FB_ProductionTank
END_ACTION

ACTION act_Call_For_HMI:


g_HMI.stT91_Sens:=g_Data.stTanksSens[E_Tank_Name.T91];
g_HMI.stT92_Sens:=g_Data.stTanksSens[E_Tank_Name.T92];
g_HMI.stT93_Sens:=g_Data.stTanksSens[E_Tank_Name.T93];
g_HMI.stT94_Sens:=g_Data.stTanksSens[E_Tank_Name.T94];

g_HMI.stT1_Sens:=g_Data.stTanksSens[E_Tank_Name.T1];
g_HMI.stT2_Sens:=g_Data.stTanksSens[E_Tank_Name.T2];
g_HMI.stT3_Sens:=g_Data.stTanksSens[E_Tank_Name.T3];
g_HMI.stT4_Sens:=g_Data.stTanksSens[E_Tank_Name.T4];
END_ACTION

ACTION act_Call_ProcessCntrl:
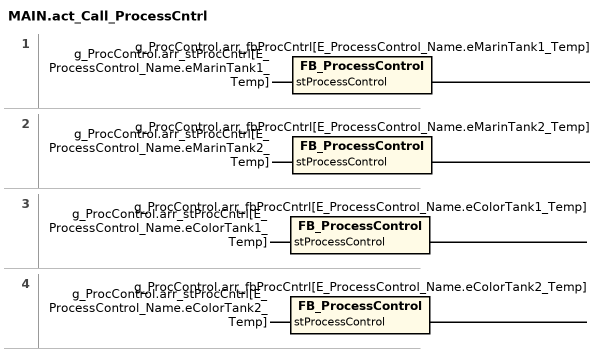
// NETWORK 1
g_ProcControl.arr_fbProcCntrl[E_ProcessControl_Name.eMarinTank1_Temp](stProcessControl := g_ProcControl.arr_stProcCntrl[E_ProcessControl_Name.eMarinTank1_Temp]); // FB_ProcessControl

// NETWORK 2
g_ProcControl.arr_fbProcCntrl[E_ProcessControl_Name.eMarinTank2_Temp](stProcessControl := g_ProcControl.arr_stProcCntrl[E_ProcessControl_Name.eMarinTank2_Temp]); // FB_ProcessControl

// NETWORK 3
g_ProcControl.arr_fbProcCntrl[E_ProcessControl_Name.eColorTank1_Temp](stProcessControl := g_ProcControl.arr_stProcCntrl[E_ProcessControl_Name.eColorTank1_Temp]); // FB_ProcessControl

// NETWORK 4
g_ProcControl.arr_fbProcCntrl[E_ProcessControl_Name.eColorTank2_Temp](stProcessControl := g_ProcControl.arr_stProcCntrl[E_ProcessControl_Name.eColorTank2_Temp]); // FB_ProcessControl
END_ACTION

ACTION act_Call_Production:

g_Prod.fbProdRecipe_Manage();
END_ACTION

ACTION act_Call_Pump_TB:
IF fbElement[E_Element_List.eTriBlender_Color].m_Get_InterConnection()=E_InterConnection.ConnToCIP 
OR fbElement[E_Element_List.eTriBlender_Marinada].m_Get_InterConnection()=E_InterConnection.ConnToCIP 
OR FALSE
THEN;
	act_Call_Pump_TB_CIP();
ELSE;
	CASE g_Data.eTriBlenderUsage OF
		E_TriBlenderUsage.eMarinada_T1,E_TriBlenderUsage.eMarinada_T2:;
				act_Call_Pump_TB_M();
		E_TriBlenderUsage.eColor_T3,E_TriBlenderUsage.eColor_T4:;
				act_Call_Pump_TB_C();
	ELSE;
		act_Call_Pump_TB_0();
	END_CASE	
END_IF
END_ACTION

ACTION act_Call_Pump_TB_0:
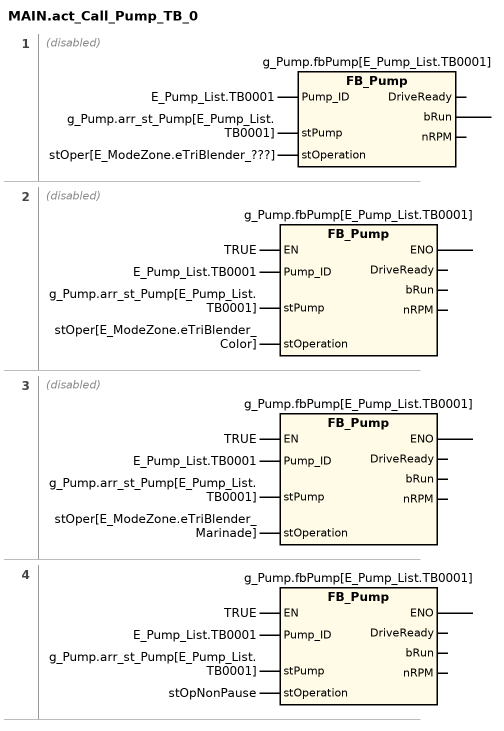
// NETWORK 1 (disabled)
// g_Pump.fbPump[E_Pump_List.TB0001](
//     Pump_ID := E_Pump_List.TB0001,
//     stPump := g_Pump.arr_st_Pump[E_Pump_List.TB0001],
//     stOperation := stOper[E_ModeZone.eTriBlender_???]); // FB_Pump

// NETWORK 2 (disabled)
// g_Pump.fbPump[E_Pump_List.TB0001](
//     Pump_ID := E_Pump_List.TB0001,
//     stPump := g_Pump.arr_st_Pump[E_Pump_List.TB0001],
//     stOperation := stOper[E_ModeZone.eTriBlender_Color]); // FB_Pump

// NETWORK 3 (disabled)
// g_Pump.fbPump[E_Pump_List.TB0001](
//     Pump_ID := E_Pump_List.TB0001,
//     stPump := g_Pump.arr_st_Pump[E_Pump_List.TB0001],
//     stOperation := stOper[E_ModeZone.eTriBlender_Marinade]); // FB_Pump

// NETWORK 4
g_Pump.fbPump[E_Pump_List.TB0001](
    Pump_ID := E_Pump_List.TB0001,
    stPump := g_Pump.arr_st_Pump[E_Pump_List.TB0001],
    stOperation := stOpNonPause); // FB_Pump
END_ACTION

ACTION act_Call_Pump_TB_C:
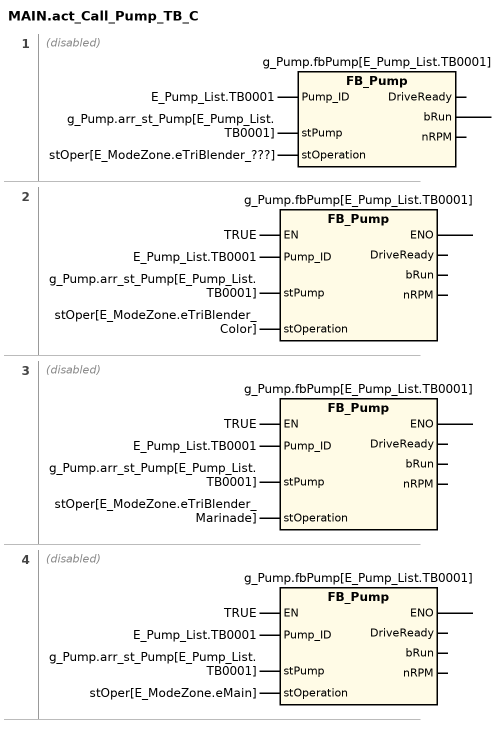
// NETWORK 1 (disabled)
// g_Pump.fbPump[E_Pump_List.TB0001](
//     Pump_ID := E_Pump_List.TB0001,
//     stPump := g_Pump.arr_st_Pump[E_Pump_List.TB0001],
//     stOperation := stOper[E_ModeZone.eTriBlender_???]); // FB_Pump

// NETWORK 2
g_Pump.fbPump[E_Pump_List.TB0001](
    Pump_ID := E_Pump_List.TB0001,
    stPump := g_Pump.arr_st_Pump[E_Pump_List.TB0001],
    stOperation := stOper[E_ModeZone.eTriBlender_Color]); // FB_Pump

// NETWORK 3 (disabled)
// g_Pump.fbPump[E_Pump_List.TB0001](
//     Pump_ID := E_Pump_List.TB0001,
//     stPump := g_Pump.arr_st_Pump[E_Pump_List.TB0001],
//     stOperation := stOper[E_ModeZone.eTriBlender_Marinade]); // FB_Pump

// NETWORK 4 (disabled)
// g_Pump.fbPump[E_Pump_List.TB0001](
//     Pump_ID := E_Pump_List.TB0001,
//     stPump := g_Pump.arr_st_Pump[E_Pump_List.TB0001],
//     stOperation := stOper[E_ModeZone.eMain]); // FB_Pump
END_ACTION

ACTION act_Call_Pump_TB_CIP:
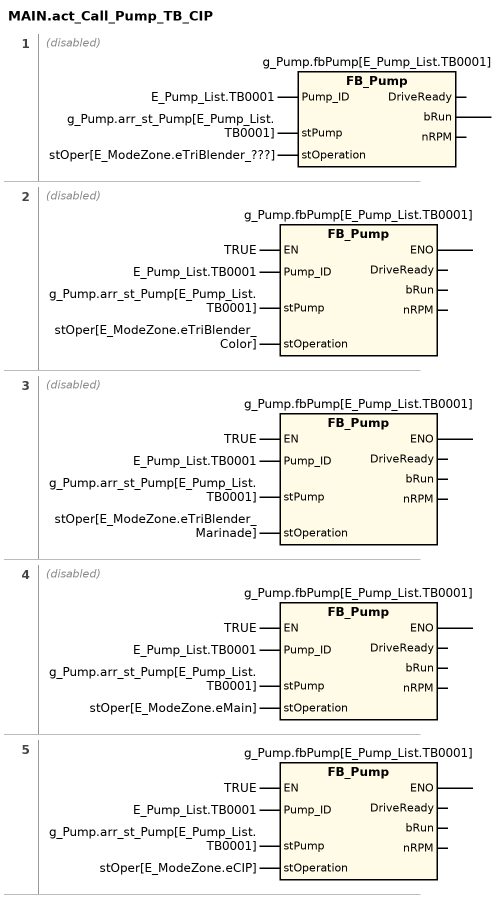
// NETWORK 1 (disabled)
// g_Pump.fbPump[E_Pump_List.TB0001](
//     Pump_ID := E_Pump_List.TB0001,
//     stPump := g_Pump.arr_st_Pump[E_Pump_List.TB0001],
//     stOperation := stOper[E_ModeZone.eTriBlender_???]); // FB_Pump

// NETWORK 2 (disabled)
// g_Pump.fbPump[E_Pump_List.TB0001](
//     Pump_ID := E_Pump_List.TB0001,
//     stPump := g_Pump.arr_st_Pump[E_Pump_List.TB0001],
//     stOperation := stOper[E_ModeZone.eTriBlender_Color]); // FB_Pump

// NETWORK 3 (disabled)
// g_Pump.fbPump[E_Pump_List.TB0001](
//     Pump_ID := E_Pump_List.TB0001,
//     stPump := g_Pump.arr_st_Pump[E_Pump_List.TB0001],
//     stOperation := stOper[E_ModeZone.eTriBlender_Marinade]); // FB_Pump

// NETWORK 4 (disabled)
// g_Pump.fbPump[E_Pump_List.TB0001](
//     Pump_ID := E_Pump_List.TB0001,
//     stPump := g_Pump.arr_st_Pump[E_Pump_List.TB0001],
//     stOperation := stOper[E_ModeZone.eMain]); // FB_Pump

// NETWORK 5
g_Pump.fbPump[E_Pump_List.TB0001](
    Pump_ID := E_Pump_List.TB0001,
    stPump := g_Pump.arr_st_Pump[E_Pump_List.TB0001],
    stOperation := stOper[E_ModeZone.eCIP]); // FB_Pump
END_ACTION

ACTION act_Call_Pump_TB_M:
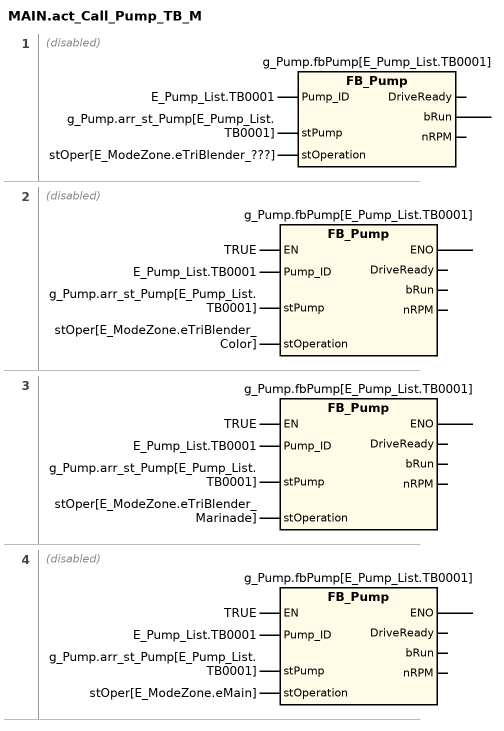
// NETWORK 1 (disabled)
// g_Pump.fbPump[E_Pump_List.TB0001](
//     Pump_ID := E_Pump_List.TB0001,
//     stPump := g_Pump.arr_st_Pump[E_Pump_List.TB0001],
//     stOperation := stOper[E_ModeZone.eTriBlender_???]); // FB_Pump

// NETWORK 2 (disabled)
// g_Pump.fbPump[E_Pump_List.TB0001](
//     Pump_ID := E_Pump_List.TB0001,
//     stPump := g_Pump.arr_st_Pump[E_Pump_List.TB0001],
//     stOperation := stOper[E_ModeZone.eTriBlender_Color]); // FB_Pump

// NETWORK 3
g_Pump.fbPump[E_Pump_List.TB0001](
    Pump_ID := E_Pump_List.TB0001,
    stPump := g_Pump.arr_st_Pump[E_Pump_List.TB0001],
    stOperation := stOper[E_ModeZone.eTriBlender_Marinade]); // FB_Pump

// NETWORK 4 (disabled)
// g_Pump.fbPump[E_Pump_List.TB0001](
//     Pump_ID := E_Pump_List.TB0001,
//     stPump := g_Pump.arr_st_Pump[E_Pump_List.TB0001],
//     stOperation := stOper[E_ModeZone.eMain]); // FB_Pump
END_ACTION

ACTION act_Call_Pumps:
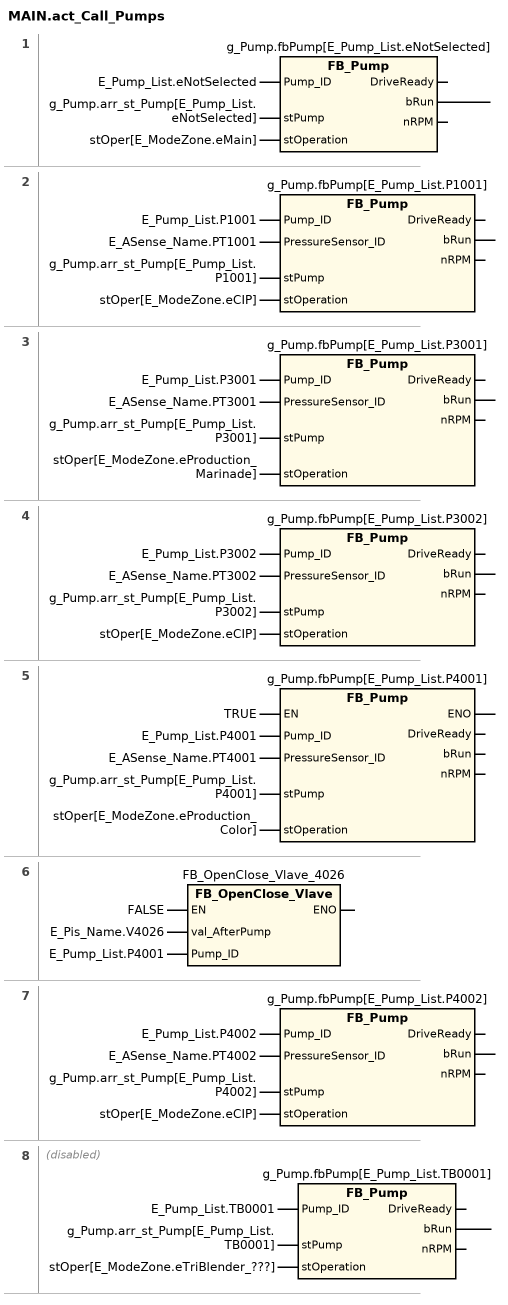
// NETWORK 1
g_Pump.fbPump[E_Pump_List.eNotSelected](
    Pump_ID := E_Pump_List.eNotSelected,
    stPump := g_Pump.arr_st_Pump[E_Pump_List.eNotSelected],
    stOperation := stOper[E_ModeZone.eMain]); // FB_Pump

// NETWORK 2
g_Pump.fbPump[E_Pump_List.P1001](
    Pump_ID := E_Pump_List.P1001,
    PressureSensor_ID := E_ASense_Name.PT1001,
    stPump := g_Pump.arr_st_Pump[E_Pump_List.P1001],
    stOperation := stOper[E_ModeZone.eCIP]); // FB_Pump

// NETWORK 3
g_Pump.fbPump[E_Pump_List.P3001](
    Pump_ID := E_Pump_List.P3001,
    PressureSensor_ID := E_ASense_Name.PT3001,
    stPump := g_Pump.arr_st_Pump[E_Pump_List.P3001],
    stOperation := stOper[E_ModeZone.eProduction_Marinade]); // FB_Pump

// NETWORK 4
g_Pump.fbPump[E_Pump_List.P3002](
    Pump_ID := E_Pump_List.P3002,
    PressureSensor_ID := E_ASense_Name.PT3002,
    stPump := g_Pump.arr_st_Pump[E_Pump_List.P3002],
    stOperation := stOper[E_ModeZone.eCIP]); // FB_Pump

// NETWORK 5
g_Pump.fbPump[E_Pump_List.P4001](
    Pump_ID := E_Pump_List.P4001,
    PressureSensor_ID := E_ASense_Name.PT4001,
    stPump := g_Pump.arr_st_Pump[E_Pump_List.P4001],
    stOperation := stOper[E_ModeZone.eProduction_Color]); // FB_Pump

// NETWORK 6
IF FALSE THEN
    FB_OpenClose_Vlave_4026(val_AfterPump := E_Pis_Name.V4026, Pump_ID := E_Pump_List.P4001); // FB_OpenClose_Vlave
END_IF

// NETWORK 7
g_Pump.fbPump[E_Pump_List.P4002](
    Pump_ID := E_Pump_List.P4002,
    PressureSensor_ID := E_ASense_Name.PT4002,
    stPump := g_Pump.arr_st_Pump[E_Pump_List.P4002],
    stOperation := stOper[E_ModeZone.eCIP]); // FB_Pump

// NETWORK 8 (disabled)
// g_Pump.fbPump[E_Pump_List.TB0001](
//     Pump_ID := E_Pump_List.TB0001,
//     stPump := g_Pump.arr_st_Pump[E_Pump_List.TB0001],
//     stOperation := stOper[E_ModeZone.eTriBlender_???]); // FB_Pump

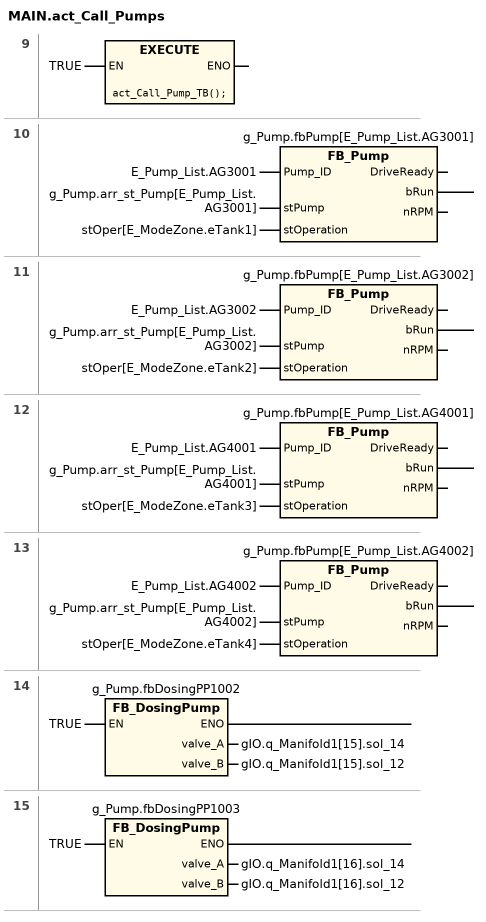
// NETWORK 9

act_Call_Pump_TB();

// NETWORK 10
g_Pump.fbPump[E_Pump_List.AG3001](
    Pump_ID := E_Pump_List.AG3001,
    stPump := g_Pump.arr_st_Pump[E_Pump_List.AG3001],
    stOperation := stOper[E_ModeZone.eTank1]); // FB_Pump

// NETWORK 11
g_Pump.fbPump[E_Pump_List.AG3002](
    Pump_ID := E_Pump_List.AG3002,
    stPump := g_Pump.arr_st_Pump[E_Pump_List.AG3002],
    stOperation := stOper[E_ModeZone.eTank2]); // FB_Pump

// NETWORK 12
g_Pump.fbPump[E_Pump_List.AG4001](
    Pump_ID := E_Pump_List.AG4001,
    stPump := g_Pump.arr_st_Pump[E_Pump_List.AG4001],
    stOperation := stOper[E_ModeZone.eTank3]); // FB_Pump

// NETWORK 13
g_Pump.fbPump[E_Pump_List.AG4002](
    Pump_ID := E_Pump_List.AG4002,
    stPump := g_Pump.arr_st_Pump[E_Pump_List.AG4002],
    stOperation := stOper[E_ModeZone.eTank4]); // FB_Pump

// NETWORK 14
g_Pump.fbDosingPP1002(valve_A => gIO.q_Manifold1[15].sol_14, valve_B => gIO.q_Manifold1[15].sol_12); // FB_DosingPump

// NETWORK 15
g_Pump.fbDosingPP1003(valve_A => gIO.q_Manifold1[16].sol_14, valve_B => gIO.q_Manifold1[16].sol_12); // FB_DosingPump
END_ACTION

ACTION act_Call_ScaleFactor:
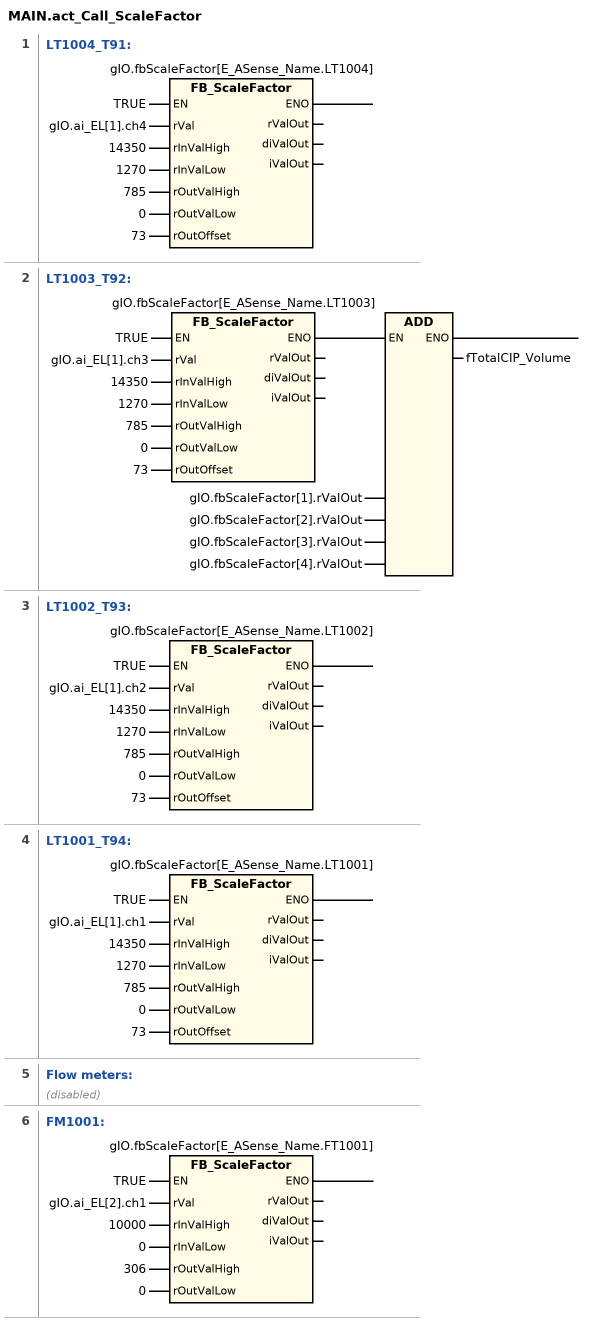
// NETWORK 1
LT1004_T91:
gIO.fbScaleFactor[E_ASense_Name.LT1004](
    rVal := gIO.ai_EL[1].ch4,
    rInValHigh := 14350,
    rInValLow := 1270,
    rOutValHigh := 785,
    rOutValLow := 0,
    rOutOffset := 73); // FB_ScaleFactor

// NETWORK 2
LT1003_T92:
gIO.fbScaleFactor[E_ASense_Name.LT1003](
    rVal := gIO.ai_EL[1].ch3,
    rInValHigh := 14350,
    rInValLow := 1270,
    rOutValHigh := 785,
    rOutValLow := 0,
    rOutOffset := 73); // FB_ScaleFactor
fTotalCIP_Volume := gIO.fbScaleFactor[1].rValOut + gIO.fbScaleFactor[2].rValOut + gIO.fbScaleFactor[3].rValOut + gIO.fbScaleFactor[4].rValOut;

// NETWORK 3
LT1002_T93:
gIO.fbScaleFactor[E_ASense_Name.LT1002](
    rVal := gIO.ai_EL[1].ch2,
    rInValHigh := 14350,
    rInValLow := 1270,
    rOutValHigh := 785,
    rOutValLow := 0,
    rOutOffset := 73); // FB_ScaleFactor

// NETWORK 4
LT1001_T94:
gIO.fbScaleFactor[E_ASense_Name.LT1001](
    rVal := gIO.ai_EL[1].ch1,
    rInValHigh := 14350,
    rInValLow := 1270,
    rOutValHigh := 785,
    rOutValLow := 0,
    rOutOffset := 73); // FB_ScaleFactor

// NETWORK 5 (disabled)
// label: Flow meters

// NETWORK 6
FM1001:
gIO.fbScaleFactor[E_ASense_Name.FT1001](
    rVal := gIO.ai_EL[2].ch1,
    rInValHigh := 10000,
    rInValLow := 0,
    rOutValHigh := 306,
    rOutValLow := 0); // FB_ScaleFactor

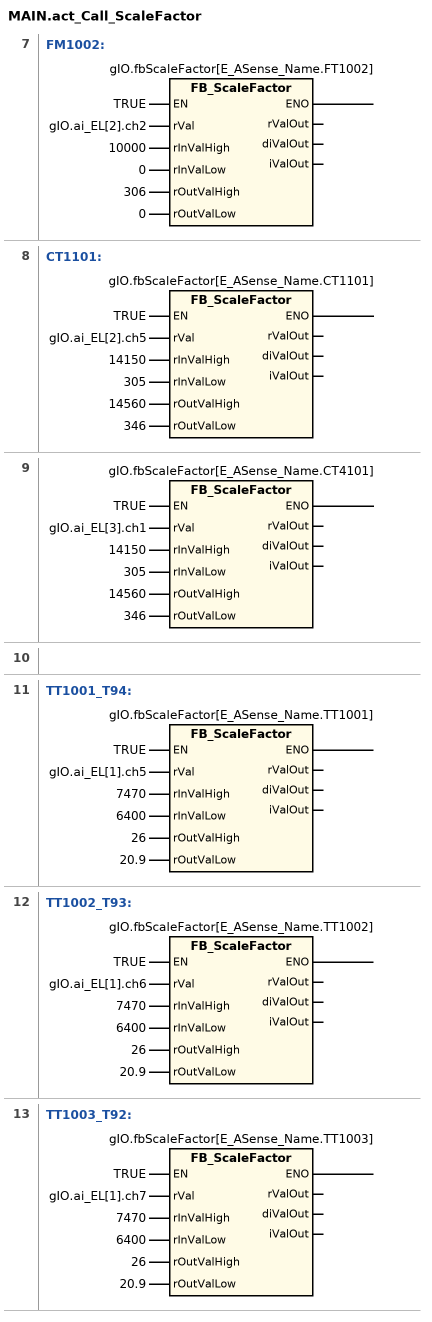
// NETWORK 7
FM1002:
gIO.fbScaleFactor[E_ASense_Name.FT1002](
    rVal := gIO.ai_EL[2].ch2,
    rInValHigh := 10000,
    rInValLow := 0,
    rOutValHigh := 306,
    rOutValLow := 0); // FB_ScaleFactor

// NETWORK 8
CT1101:
gIO.fbScaleFactor[E_ASense_Name.CT1101](
    rVal := gIO.ai_EL[2].ch5,
    rInValHigh := 14150,
    rInValLow := 305,
    rOutValHigh := 14560,
    rOutValLow := 346); // FB_ScaleFactor

// NETWORK 9
gIO.fbScaleFactor[E_ASense_Name.CT4101](
    rVal := gIO.ai_EL[3].ch1,
    rInValHigh := 14150,
    rInValLow := 305,
    rOutValHigh := 14560,
    rOutValLow := 346); // FB_ScaleFactor

// NETWORK 10

// NETWORK 11
TT1001_T94:
gIO.fbScaleFactor[E_ASense_Name.TT1001](
    rVal := gIO.ai_EL[1].ch5,
    rInValHigh := 7470,
    rInValLow := 6400,
    rOutValHigh := 26,
    rOutValLow := 20.9); // FB_ScaleFactor

// NETWORK 12
TT1002_T93:
gIO.fbScaleFactor[E_ASense_Name.TT1002](
    rVal := gIO.ai_EL[1].ch6,
    rInValHigh := 7470,
    rInValLow := 6400,
    rOutValHigh := 26,
    rOutValLow := 20.9); // FB_ScaleFactor

// NETWORK 13
TT1003_T92:
gIO.fbScaleFactor[E_ASense_Name.TT1003](
    rVal := gIO.ai_EL[1].ch7,
    rInValHigh := 7470,
    rInValLow := 6400,
    rOutValHigh := 26,
    rOutValLow := 20.9); // FB_ScaleFactor

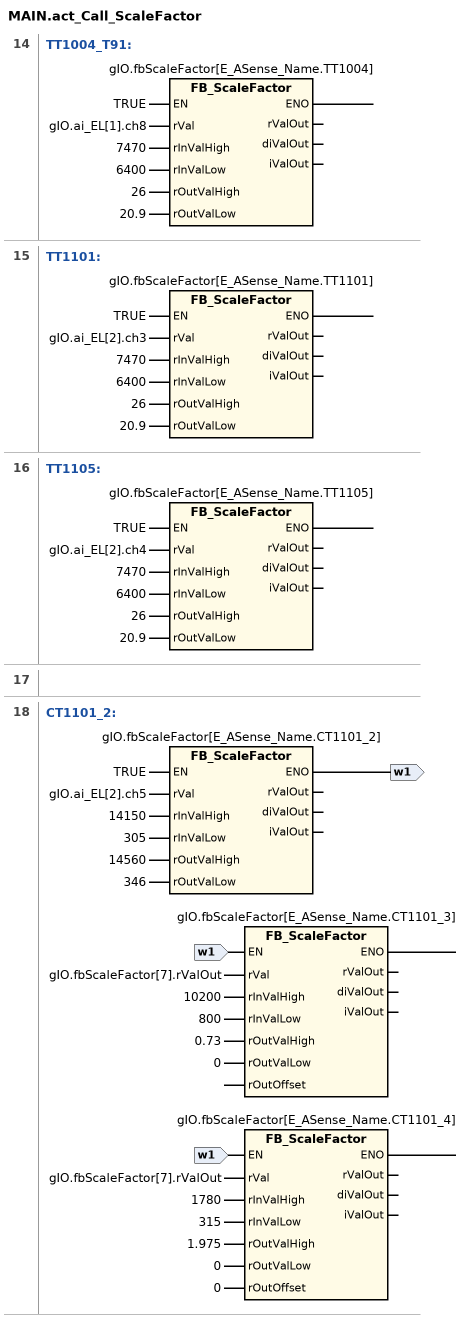
// NETWORK 14
TT1004_T91:
gIO.fbScaleFactor[E_ASense_Name.TT1004](
    rVal := gIO.ai_EL[1].ch8,
    rInValHigh := 7470,
    rInValLow := 6400,
    rOutValHigh := 26,
    rOutValLow := 20.9); // FB_ScaleFactor

// NETWORK 15
TT1101:
gIO.fbScaleFactor[E_ASense_Name.TT1101](
    rVal := gIO.ai_EL[2].ch3,
    rInValHigh := 7470,
    rInValLow := 6400,
    rOutValHigh := 26,
    rOutValLow := 20.9); // FB_ScaleFactor

// NETWORK 16
TT1105:
gIO.fbScaleFactor[E_ASense_Name.TT1105](
    rVal := gIO.ai_EL[2].ch4,
    rInValHigh := 7470,
    rInValLow := 6400,
    rOutValHigh := 26,
    rOutValLow := 20.9); // FB_ScaleFactor

// NETWORK 17

// NETWORK 18
CT1101_2:
gIO.fbScaleFactor[E_ASense_Name.CT1101_2](
    rVal := gIO.ai_EL[2].ch5,
    rInValHigh := 14150,
    rInValLow := 305,
    rOutValHigh := 14560,
    rOutValLow := 346); // FB_ScaleFactor
gIO.fbScaleFactor[E_ASense_Name.CT1101_3](
    rVal := gIO.fbScaleFactor[7].rValOut,
    rInValHigh := 10200,
    rInValLow := 800,
    rOutValHigh := 0.73,
    rOutValLow := 0); // FB_ScaleFactor
gIO.fbScaleFactor[E_ASense_Name.CT1101_4](
    rVal := gIO.fbScaleFactor[7].rValOut,
    rInValHigh := 1780,
    rInValLow := 315,
    rOutValHigh := 1.975,
    rOutValLow := 0,
    rOutOffset := 0); // FB_ScaleFactor

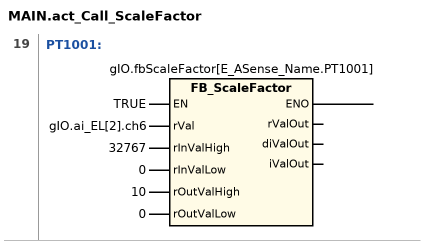
// NETWORK 19
PT1001:
gIO.fbScaleFactor[E_ASense_Name.PT1001](
    rVal := gIO.ai_EL[2].ch6,
    rInValHigh := 32767,
    rInValLow := 0,
    rOutValHigh := 10,
    rOutValLow := 0); // FB_ScaleFactor
END_ACTION

ACTION act_Call_Sensors_Analog:
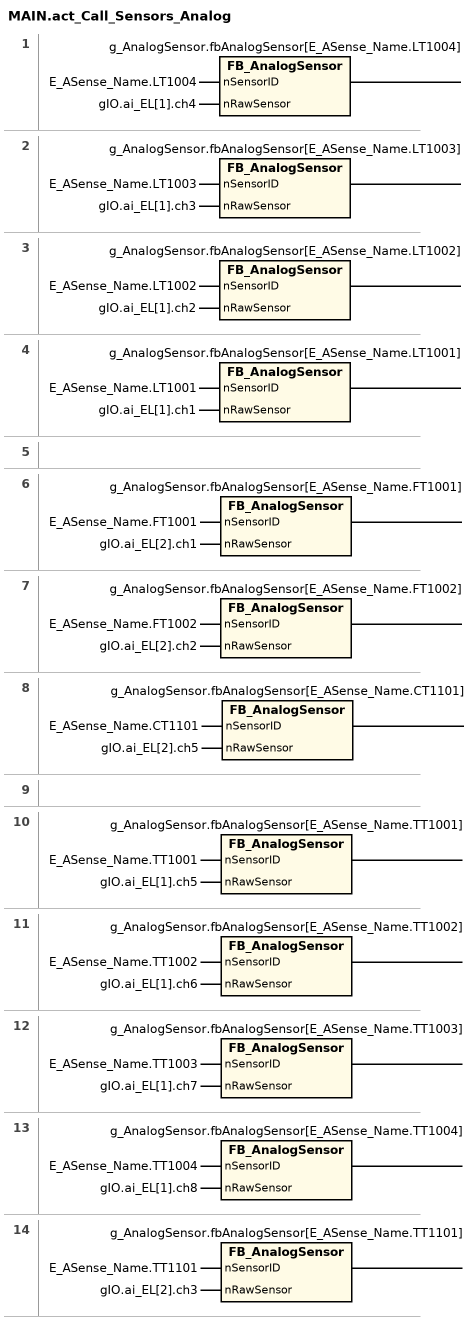
// NETWORK 1
g_AnalogSensor.fbAnalogSensor[E_ASense_Name.LT1004](nSensorID := E_ASense_Name.LT1004, nRawSensor := gIO.ai_EL[1].ch4); // FB_AnalogSensor

// NETWORK 2
g_AnalogSensor.fbAnalogSensor[E_ASense_Name.LT1003](nSensorID := E_ASense_Name.LT1003, nRawSensor := gIO.ai_EL[1].ch3); // FB_AnalogSensor

// NETWORK 3
g_AnalogSensor.fbAnalogSensor[E_ASense_Name.LT1002](nSensorID := E_ASense_Name.LT1002, nRawSensor := gIO.ai_EL[1].ch2); // FB_AnalogSensor

// NETWORK 4
g_AnalogSensor.fbAnalogSensor[E_ASense_Name.LT1001](nSensorID := E_ASense_Name.LT1001, nRawSensor := gIO.ai_EL[1].ch1); // FB_AnalogSensor

// NETWORK 5

// NETWORK 6
g_AnalogSensor.fbAnalogSensor[E_ASense_Name.FT1001](nSensorID := E_ASense_Name.FT1001, nRawSensor := gIO.ai_EL[2].ch1); // FB_AnalogSensor

// NETWORK 7
g_AnalogSensor.fbAnalogSensor[E_ASense_Name.FT1002](nSensorID := E_ASense_Name.FT1002, nRawSensor := gIO.ai_EL[2].ch2); // FB_AnalogSensor

// NETWORK 8
g_AnalogSensor.fbAnalogSensor[E_ASense_Name.CT1101](nSensorID := E_ASense_Name.CT1101, nRawSensor := gIO.ai_EL[2].ch5); // FB_AnalogSensor

// NETWORK 9

// NETWORK 10
g_AnalogSensor.fbAnalogSensor[E_ASense_Name.TT1001](nSensorID := E_ASense_Name.TT1001, nRawSensor := gIO.ai_EL[1].ch5); // FB_AnalogSensor

// NETWORK 11
g_AnalogSensor.fbAnalogSensor[E_ASense_Name.TT1002](nSensorID := E_ASense_Name.TT1002, nRawSensor := gIO.ai_EL[1].ch6); // FB_AnalogSensor

// NETWORK 12
g_AnalogSensor.fbAnalogSensor[E_ASense_Name.TT1003](nSensorID := E_ASense_Name.TT1003, nRawSensor := gIO.ai_EL[1].ch7); // FB_AnalogSensor

// NETWORK 13
g_AnalogSensor.fbAnalogSensor[E_ASense_Name.TT1004](nSensorID := E_ASense_Name.TT1004, nRawSensor := gIO.ai_EL[1].ch8); // FB_AnalogSensor

// NETWORK 14
g_AnalogSensor.fbAnalogSensor[E_ASense_Name.TT1101](nSensorID := E_ASense_Name.TT1101, nRawSensor := gIO.ai_EL[2].ch3); // FB_AnalogSensor

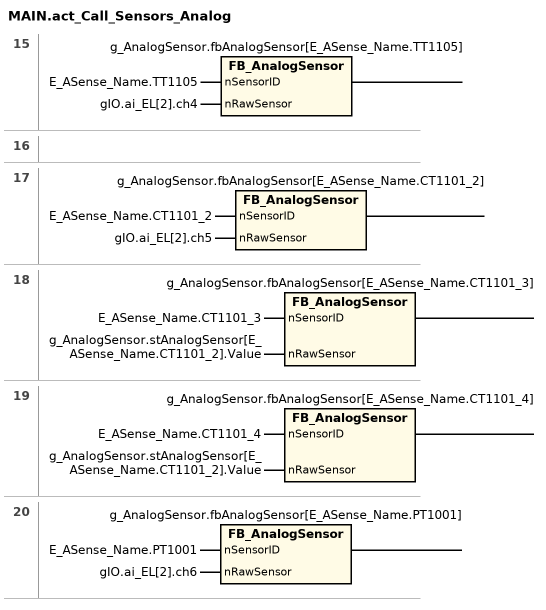
// NETWORK 15
g_AnalogSensor.fbAnalogSensor[E_ASense_Name.TT1105](nSensorID := E_ASense_Name.TT1105, nRawSensor := gIO.ai_EL[2].ch4); // FB_AnalogSensor

// NETWORK 16

// NETWORK 17
g_AnalogSensor.fbAnalogSensor[E_ASense_Name.CT1101_2](nSensorID := E_ASense_Name.CT1101_2, nRawSensor := gIO.ai_EL[2].ch5); // FB_AnalogSensor

// NETWORK 18
g_AnalogSensor.fbAnalogSensor[E_ASense_Name.CT1101_3](nSensorID := E_ASense_Name.CT1101_3, nRawSensor := g_AnalogSensor.stAnalogSensor[E_ASense_Name.CT1101_2].Value); // FB_AnalogSensor

// NETWORK 19
g_AnalogSensor.fbAnalogSensor[E_ASense_Name.CT1101_4](nSensorID := E_ASense_Name.CT1101_4, nRawSensor := g_AnalogSensor.stAnalogSensor[E_ASense_Name.CT1101_2].Value); // FB_AnalogSensor

// NETWORK 20
g_AnalogSensor.fbAnalogSensor[E_ASense_Name.PT1001](nSensorID := E_ASense_Name.PT1001, nRawSensor := gIO.ai_EL[2].ch6); // FB_AnalogSensor
END_ACTION

ACTION act_Call_Sensors_Analog_1:
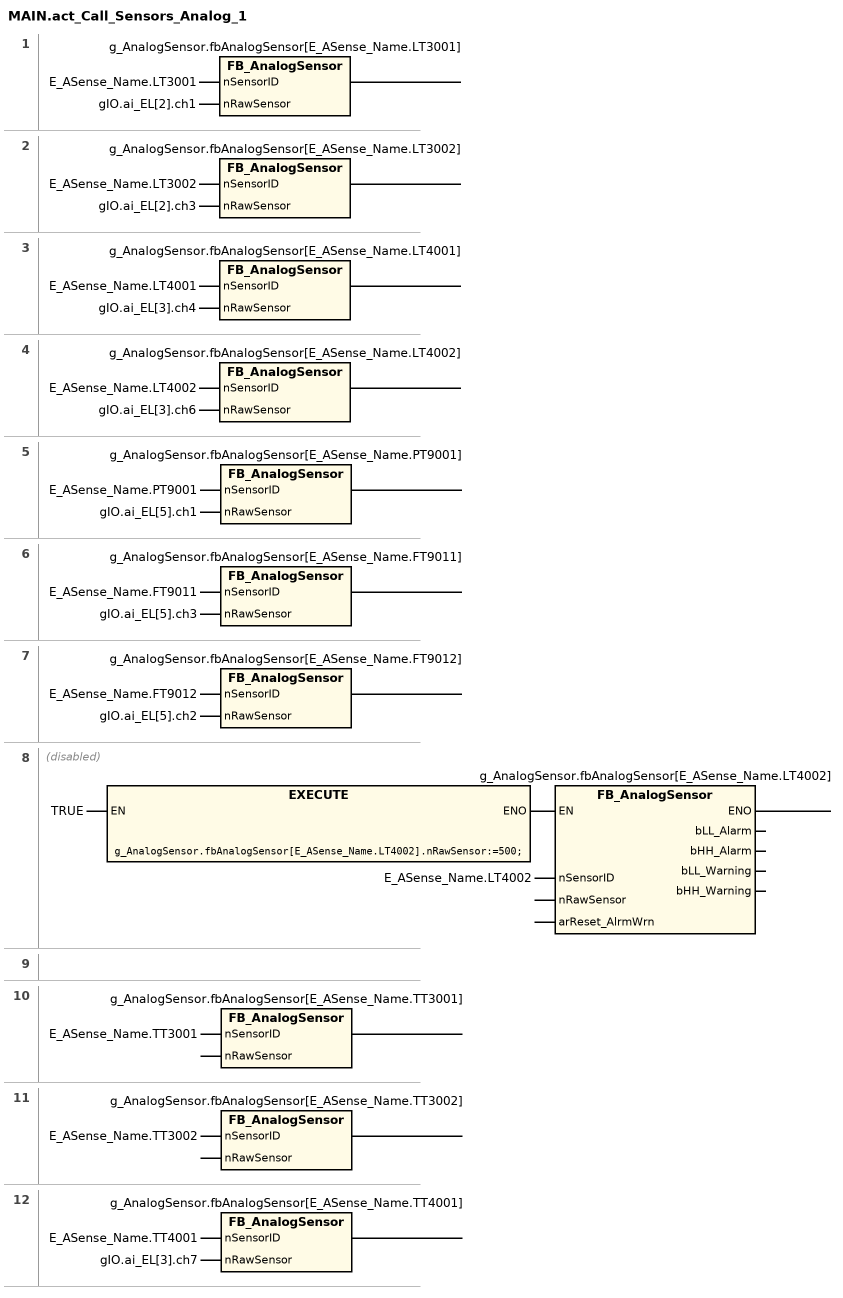
// NETWORK 1
g_AnalogSensor.fbAnalogSensor[E_ASense_Name.LT3001](nSensorID := E_ASense_Name.LT3001, nRawSensor := gIO.ai_EL[2].ch1); // FB_AnalogSensor

// NETWORK 2
g_AnalogSensor.fbAnalogSensor[E_ASense_Name.LT3002](nSensorID := E_ASense_Name.LT3002, nRawSensor := gIO.ai_EL[2].ch3); // FB_AnalogSensor

// NETWORK 3
g_AnalogSensor.fbAnalogSensor[E_ASense_Name.LT4001](nSensorID := E_ASense_Name.LT4001, nRawSensor := gIO.ai_EL[3].ch4); // FB_AnalogSensor

// NETWORK 4
g_AnalogSensor.fbAnalogSensor[E_ASense_Name.LT4002](nSensorID := E_ASense_Name.LT4002, nRawSensor := gIO.ai_EL[3].ch6); // FB_AnalogSensor

// NETWORK 5
g_AnalogSensor.fbAnalogSensor[E_ASense_Name.PT9001](nSensorID := E_ASense_Name.PT9001, nRawSensor := gIO.ai_EL[5].ch1); // FB_AnalogSensor

// NETWORK 6
g_AnalogSensor.fbAnalogSensor[E_ASense_Name.FT9011](nSensorID := E_ASense_Name.FT9011, nRawSensor := gIO.ai_EL[5].ch3); // FB_AnalogSensor

// NETWORK 7
g_AnalogSensor.fbAnalogSensor[E_ASense_Name.FT9012](nSensorID := E_ASense_Name.FT9012, nRawSensor := gIO.ai_EL[5].ch2); // FB_AnalogSensor

// NETWORK 8 (disabled)
// 
// 
// g_AnalogSensor.fbAnalogSensor[E_ASense_Name.LT4002].nRawSensor:=500;
// g_AnalogSensor.fbAnalogSensor[E_ASense_Name.LT4002](nSensorID := E_ASense_Name.LT4002); // FB_AnalogSensor

// NETWORK 9

// NETWORK 10
g_AnalogSensor.fbAnalogSensor[E_ASense_Name.TT3001](nSensorID := E_ASense_Name.TT3001); // FB_AnalogSensor

// NETWORK 11
g_AnalogSensor.fbAnalogSensor[E_ASense_Name.TT3002](nSensorID := E_ASense_Name.TT3002); // FB_AnalogSensor

// NETWORK 12
g_AnalogSensor.fbAnalogSensor[E_ASense_Name.TT4001](nSensorID := E_ASense_Name.TT4001, nRawSensor := gIO.ai_EL[3].ch7); // FB_AnalogSensor

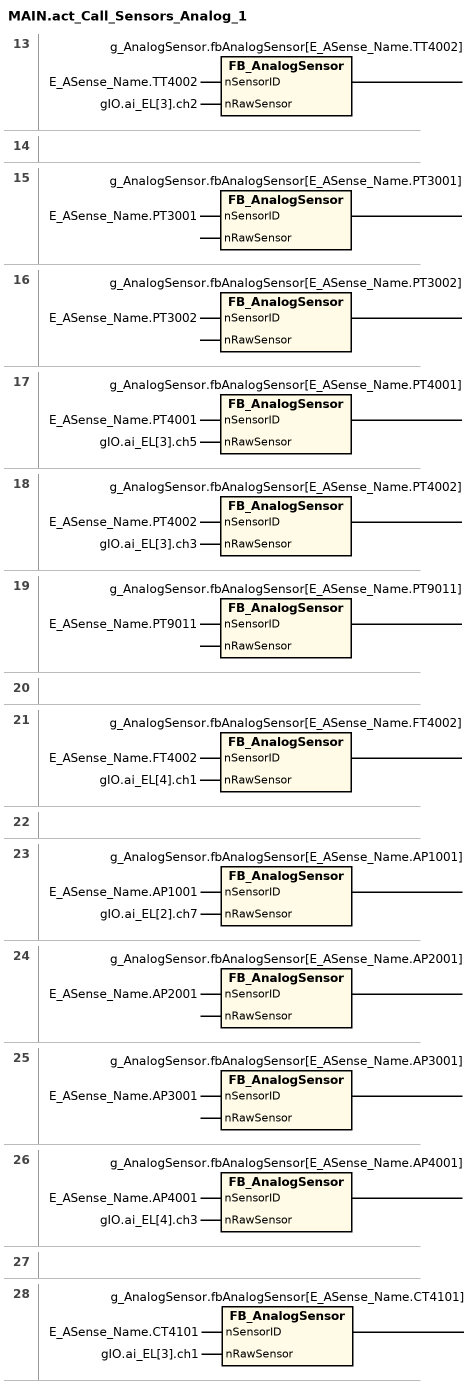
// NETWORK 13
g_AnalogSensor.fbAnalogSensor[E_ASense_Name.TT4002](nSensorID := E_ASense_Name.TT4002, nRawSensor := gIO.ai_EL[3].ch2); // FB_AnalogSensor

// NETWORK 14

// NETWORK 15
g_AnalogSensor.fbAnalogSensor[E_ASense_Name.PT3001](nSensorID := E_ASense_Name.PT3001); // FB_AnalogSensor

// NETWORK 16
g_AnalogSensor.fbAnalogSensor[E_ASense_Name.PT3002](nSensorID := E_ASense_Name.PT3002); // FB_AnalogSensor

// NETWORK 17
g_AnalogSensor.fbAnalogSensor[E_ASense_Name.PT4001](nSensorID := E_ASense_Name.PT4001, nRawSensor := gIO.ai_EL[3].ch5); // FB_AnalogSensor

// NETWORK 18
g_AnalogSensor.fbAnalogSensor[E_ASense_Name.PT4002](nSensorID := E_ASense_Name.PT4002, nRawSensor := gIO.ai_EL[3].ch3); // FB_AnalogSensor

// NETWORK 19
g_AnalogSensor.fbAnalogSensor[E_ASense_Name.PT9011](nSensorID := E_ASense_Name.PT9011); // FB_AnalogSensor

// NETWORK 20

// NETWORK 21
g_AnalogSensor.fbAnalogSensor[E_ASense_Name.FT4002](nSensorID := E_ASense_Name.FT4002, nRawSensor := gIO.ai_EL[4].ch1); // FB_AnalogSensor

// NETWORK 22

// NETWORK 23
g_AnalogSensor.fbAnalogSensor[E_ASense_Name.AP1001](nSensorID := E_ASense_Name.AP1001, nRawSensor := gIO.ai_EL[2].ch7); // FB_AnalogSensor

// NETWORK 24
g_AnalogSensor.fbAnalogSensor[E_ASense_Name.AP2001](nSensorID := E_ASense_Name.AP2001); // FB_AnalogSensor

// NETWORK 25
g_AnalogSensor.fbAnalogSensor[E_ASense_Name.AP3001](nSensorID := E_ASense_Name.AP3001); // FB_AnalogSensor

// NETWORK 26
g_AnalogSensor.fbAnalogSensor[E_ASense_Name.AP4001](nSensorID := E_ASense_Name.AP4001, nRawSensor := gIO.ai_EL[4].ch3); // FB_AnalogSensor

// NETWORK 27

// NETWORK 28
g_AnalogSensor.fbAnalogSensor[E_ASense_Name.CT4101](nSensorID := E_ASense_Name.CT4101, nRawSensor := gIO.ai_EL[3].ch1); // FB_AnalogSensor

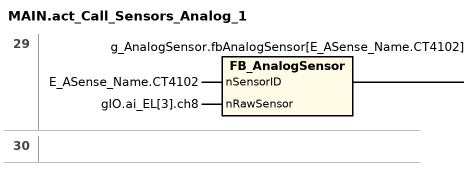
// NETWORK 29
g_AnalogSensor.fbAnalogSensor[E_ASense_Name.CT4102](nSensorID := E_ASense_Name.CT4102, nRawSensor := gIO.ai_EL[3].ch8); // FB_AnalogSensor

// NETWORK 30
END_ACTION

ACTION act_ClientPump_Select:
CASE arCIP_RequestBufer[0].eClient OF
	E_CIP_Usage.eTank_1,
	E_CIP_Usage.eTank_2:;
				eClientPump:=E_Pump_List.P3002;
	E_CIP_Usage.eTank_3,
	E_CIP_Usage.eTank_4:;
				eClientPump:=E_Pump_List.P4002;
	E_CIP_Usage.eLine_Marinada:;
				eClientPump:=E_Pump_List.P3001;
	E_CIP_Usage.eLine_Color:;
				eClientPump:=E_Pump_List.P4001;
	E_CIP_Usage.eTriBlender_Marinada,
	E_CIP_Usage.eTriBlender_Color:;
				eClientPump:=E_Pump_List.TB0001;
	E_CIP_Usage.eLocal:;
				eClientPump:=E_Pump_List.eNotSelected;
END_CASE
END_ACTION

ACTION act_ClientStirrer_Select:
CASE arCIP_RequestBufer[0].eClient OF
	E_CIP_Usage.eTank_1:;
				eClientStirrer:=E_Pump_List.AG3001;
	E_CIP_Usage.eTank_2:;
				eClientStirrer:=E_Pump_List.AG3002;
	E_CIP_Usage.eTank_3:;
				eClientStirrer:=E_Pump_List.AG4001;
	E_CIP_Usage.eTank_4:;
				eClientStirrer:=E_Pump_List.AG4002;
				
	(*E_CIP_Usage.eLine_Marinada:;
	E_CIP_Usage.eLine_Color:;
	E_CIP_Usage.eTriBlender_Marinada,
	E_CIP_Usage.eTriBlender_Color:;*)
ELSE;
	eClientStirrer:=E_Pump_List.eNotSelected;			
END_CASE
END_ACTION

ACTION act_HeatExchenger:
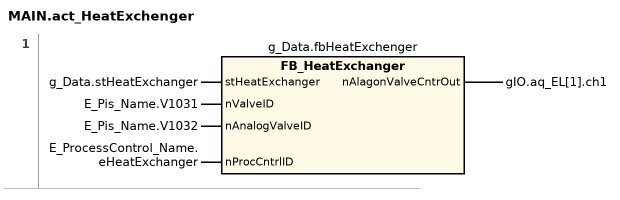
// NETWORK 1
g_Data.fbHeatExchenger(
    stHeatExchanger := g_Data.stHeatExchanger,
    nValveID := E_Pis_Name.V1031,
    nAnalogValveID := E_Pis_Name.V1032,
    nProcCntrlID := E_ProcessControl_Name.eHeatExchanger); // FB_HeatExchanger
gIO.aq_EL[1].ch1 := g_Data.fbHeatExchenger.nAlagonValveCntrOut;
END_ACTION

ACTION act_ResetPumps:
(*ftg_EStop_Fall(CLK:=prg_Safety.ftStateSafe.Q , Q=> );//EStop falling signal
rs_EStopFall(SET:=ftg_EStop_Fall.Q , RESET1:= , Q1=> );
IF rs_EStopFall.Q1 THEN
	FOR nI_1:=1 TO E_Pump_List.last BY 1 DO
		g_Pump.arr_st_Pump[nI_1].bRun_Auto:=FALSE;
	END_FOR
	rs_EStopFall.RESET1:=TRUE;
END_IF
rs_EStopFall.RESET1:=FALSE;*)
;
END_ACTION

ACTION act_Sensors:
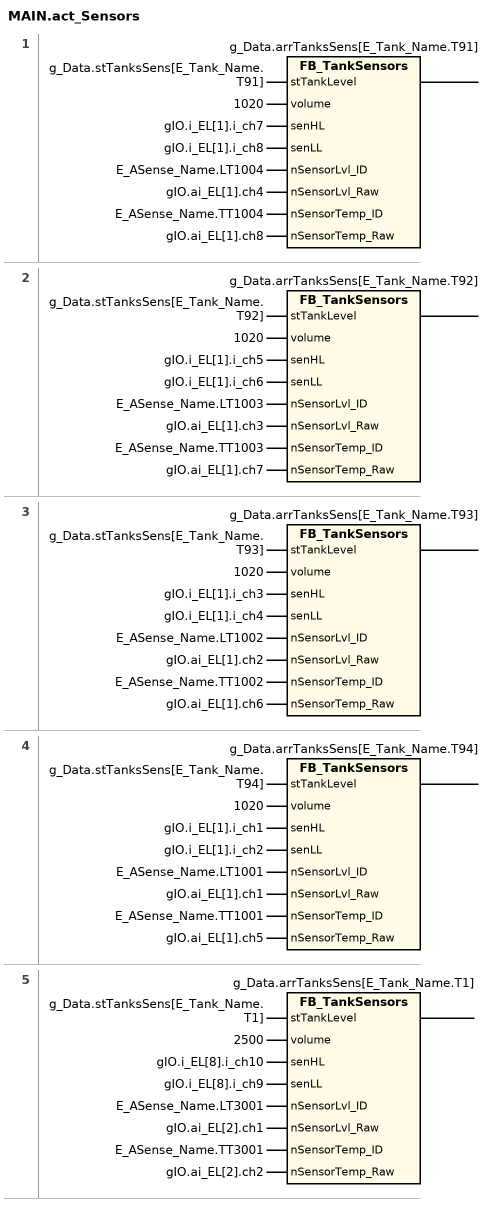
// NETWORK 1
g_Data.arrTanksSens[E_Tank_Name.T91](
    stTankLevel := g_Data.stTanksSens[E_Tank_Name.T91],
    volume := 1020,
    senHL := gIO.i_EL[1].i_ch7,
    senLL := gIO.i_EL[1].i_ch8,
    nSensorLvl_ID := E_ASense_Name.LT1004,
    nSensorLvl_Raw := gIO.ai_EL[1].ch4,
    nSensorTemp_ID := E_ASense_Name.TT1004,
    nSensorTemp_Raw := gIO.ai_EL[1].ch8); // FB_TankSensors

// NETWORK 2
g_Data.arrTanksSens[E_Tank_Name.T92](
    stTankLevel := g_Data.stTanksSens[E_Tank_Name.T92],
    volume := 1020,
    senHL := gIO.i_EL[1].i_ch5,
    senLL := gIO.i_EL[1].i_ch6,
    nSensorLvl_ID := E_ASense_Name.LT1003,
    nSensorLvl_Raw := gIO.ai_EL[1].ch3,
    nSensorTemp_ID := E_ASense_Name.TT1003,
    nSensorTemp_Raw := gIO.ai_EL[1].ch7); // FB_TankSensors

// NETWORK 3
g_Data.arrTanksSens[E_Tank_Name.T93](
    stTankLevel := g_Data.stTanksSens[E_Tank_Name.T93],
    volume := 1020,
    senHL := gIO.i_EL[1].i_ch3,
    senLL := gIO.i_EL[1].i_ch4,
    nSensorLvl_ID := E_ASense_Name.LT1002,
    nSensorLvl_Raw := gIO.ai_EL[1].ch2,
    nSensorTemp_ID := E_ASense_Name.TT1002,
    nSensorTemp_Raw := gIO.ai_EL[1].ch6); // FB_TankSensors

// NETWORK 4
g_Data.arrTanksSens[E_Tank_Name.T94](
    stTankLevel := g_Data.stTanksSens[E_Tank_Name.T94],
    volume := 1020,
    senHL := gIO.i_EL[1].i_ch1,
    senLL := gIO.i_EL[1].i_ch2,
    nSensorLvl_ID := E_ASense_Name.LT1001,
    nSensorLvl_Raw := gIO.ai_EL[1].ch1,
    nSensorTemp_ID := E_ASense_Name.TT1001,
    nSensorTemp_Raw := gIO.ai_EL[1].ch5); // FB_TankSensors

// NETWORK 5
g_Data.arrTanksSens[E_Tank_Name.T1](
    stTankLevel := g_Data.stTanksSens[E_Tank_Name.T1],
    volume := 2500,
    senHL := gIO.i_EL[8].i_ch10,
    senLL := gIO.i_EL[8].i_ch9,
    nSensorLvl_ID := E_ASense_Name.LT3001,
    nSensorLvl_Raw := gIO.ai_EL[2].ch1,
    nSensorTemp_ID := E_ASense_Name.TT3001,
    nSensorTemp_Raw := gIO.ai_EL[2].ch2); // FB_TankSensors

